(* IEC 61131-3 sources: volt/packages/volt-lsp-iec/test-corpus/awa-palletizer/Device/Plc Logic/Application/Library Manager/L_TB2P_TechModulesBasic, 108 files *)

(* ---- L_TB2P_ALLOWEDDIRECTION.dut ---- *)
TYPE L_TB2P_ALLOWEDDIRECTION :
(
	BOTH := 0,
	POSITIVE := 1,
	NEGATIVE := 2
);
END_TYPE

(* ---- L_TB2P_BASEIN.dut ---- *)
TYPE L_TB2P_BASEIN :
STRUCT
	XENABLE : BOOL;
	XRESETERROR : BOOL;
END_STRUCT
END_TYPE

(* ---- L_TB2P_BASEOUT.dut ---- *)
TYPE L_TB2P_BASEOUT :
STRUCT
	EERRORID : L_IE1P_Error;
	XWARNING : BOOL;
	XERROR : BOOL;
	ETMSTATE : L_TB2P_States := L_TB2P_States.DISABLED;
END_STRUCT
END_TYPE

(* ---- L_TB2P_BASICMOTIONBASEIN.dut ---- *)
TYPE L_TB2P_BASICMOTIONBASEIN :
STRUCT
	XUSEORIGINAL : BOOL;
	XENABLEOPERATION : BOOL;
	XQSPAPPLICATION : BOOL;
	XABORT : BOOL;
	XJOGPOS : BOOL;
	XJOGNEG : BOOL;
	XHOMEEXECUTE : BOOL;
	LROVERRIDE : LREAL := 1;
	SCCTRLBASICMOTION : L_TB2P_scCtrlBasicMotion;
END_STRUCT
END_TYPE

(* ---- L_TB2P_BASICMOTIONBASEOUT.dut ---- *)
TYPE L_TB2P_BASICMOTIONBASEOUT :
STRUCT
	XREADYFOROPERATION : BOOL;
	XOPERATIONENABLED : BOOL;
	XREADYFORMOTION : BOOL;
	XSTOACTIVE : BOOL;
	XQSPACTIVE : BOOL;
	XABORTBUSY : BOOL;
	XABORTDONE : BOOL;
	XJOGGINGBUSY : BOOL;
	XHOMINGBUSY : BOOL;
	XHOMINGDONE : BOOL;
	XISHOMED : BOOL;
	SCSTATUSBASICMOTION : L_TB2P_scStatusBasicMotion;
	LRSETACCOUT : LREAL;
	LRACTVEL : LREAL;
	LRSETVELOUT : LREAL;
	LRACTPOS : LREAL;
	LRSETPOSOUT : LREAL;
	LRACTFOLLOWINGERROR : LREAL;
END_STRUCT
END_TYPE

(* ---- L_TB2P_CATEGORY.dut ---- *)
TYPE L_TB2P_CATEGORY :
(
	DUMMY := 0
);
END_TYPE

(* ---- L_TB2P_CLASSID.dut ---- *)
TYPE L_TB2P_CLASSID :
(
	DUMMY := 0
);
END_TYPE

(* ---- L_TB2P_CLUTCHDIRECTION.dut ---- *)
TYPE L_TB2P_CLUTCHDIRECTION :
(
	MCNEGATIVEDIRECTION := -1,
	MCCURRENTDIRECTION := 0,
	MCPOSITIVEDIRECTION := 1
);
END_TYPE

(* ---- L_TB2P_CLUTCHMODE.dut ---- *)
TYPE L_TB2P_CLUTCHMODE :
(
	ABSOLUTE := 0,
	RELATIVE := 1,
	RAMP_POS := 2,
	RAMP_TIME := 3,
	DISTABSOLUTE := 4,
	ABSOLUTE_IN_TARGET := 5,
	DISTRELATIVE := 6,
	PROFGENABSOLUTE := 7,
	PROFGENRELATIVE := 8
);
END_TYPE

(* ---- L_TB2P_DIRECTION.dut ---- *)
TYPE L_TB2P_DIRECTION :
(
	BOTH := 0,
	DIRECTIONMASTER := 1
);
END_TYPE

(* ---- L_TB2P_ESELECTIONEXTTORQUELIMIT.dut ---- *)
TYPE L_TB2P_ESELECTIONEXTTORQUELIMIT :
(
	BOTHDIRECTIONS := 0,
	POSITIVEONLY := 1,
	NEGATIVEONLY := 2
);
END_TYPE

(* ---- L_TB2P_ESELECTIONMONITORINGSIGNALS.dut ---- *)
TYPE L_TB2P_ESELECTIONMONITORINGSIGNALS :
(
	NONE := 0,
	ACTUALMOTORTEMPERATURE := 1,
	ACTUALMOTORCURRENT := 2,
	DC_BUSVOLTAGE := 3,
	THERMALLOADDEVICE := 4,
	THERMALLOADMOTOR := 5,
	ANALOGSIGNAL := 6
);
END_TYPE

(* ---- L_TB2P_FBSTATES.dut ---- *)
TYPE L_TB2P_FBSTATES :
(
	INIT := 1,
	READY := 2,
	HOMING := 3,
	JOGGING := 10,
	JOGPOS := 11,
	JOGNEG := 12,
	POSITION_TRIMMING := 20,
	TRIM_POS_PLUS := 21,
	TRIM_POS_MINUS := 22,
	SYNCPOS := 30,
	POS_IS_SYNCHRONISED := 31,
	POSITIONING_TO_START_POS := 32,
	SYNCSPEED := 40,
	SPEED_IS_SYNCHRONISED := 41,
	DECOUPLED_LOCAL_DRIVING := 50,
	BASEVELOCITY := 51,
	CONTMOTION := 60,
	PREPARING_PATH := 61,
	CHECK_LIMITS := 62,
	SYNCLINEVEL := 70,
	CAMMING := 80,
	CAMMING_DONE := 81,
	CLUTCH_OPEN_INSTANT := 82,
	CLUTCH_CLOSE := 83,
	CLUTCH_OPEN := 84,
	CYCLICMOTION := 130,
	SETPARAMETERS := 140,
	CAMSEQUENCER_LOADCAMTABLE := 150,
	CAMSEQUENCER_CYCLICCAM1 := 151,
	CAMSEQUENCER_CYCLICCAM3 := 152,
	CAMSEQUENCER_CAM1CYCLICCAM3CAM1 := 153,
	CAMSEQUENCER_CAM1CAM2CYCLICCAM3CAM4CAM1 := 154,
	CALCULATION := 798,
	BUSY := 799,
	DONE := 800,
	EMERGENCYSTOP := 991,
	SLOWSTOP := 992,
	ABC := 993,
	STANDBY := 994,
	HALT := 995,
	STOP := 996,
	QUICKSTOP := 997,
	SERVICE := 998,
	ERROR := 999,
	SYSTEMFAULT := 1000
);
END_TYPE

(* ---- L_TB2P_INTERFACEID.dut ---- *)
TYPE L_TB2P_INTERFACEID :
(
	L_TB2P_ITECHMODULEBASE := (L_TB2P_Internal.cdiEnumStartValue + 1),
	L_TB2P_ITECHMODULEINTERNAL := (L_TB2P_Internal.cdiEnumStartValue + 2),
	L_TB2M_IERRORMANAGER := (L_TB2P_Internal.cdiEnumStartValue + 22),
	L_TB2P_ISTRUCTPROVIDER := (L_TB2P_Internal.cdiEnumStartValue + 23)
);
END_TYPE

(* ---- L_TB2P_SCAP_BASICMOTIONBASE.dut ---- *)
TYPE L_TB2P_SCAP_BASICMOTIONBASE :
STRUCT
END_STRUCT
END_TYPE

(* ---- L_TB2P_SCAP_TM_MOTIONCONTROL.dut ---- *)
TYPE L_TB2P_SCAP_TM_MOTIONCONTROL :
STRUCT
	AP_XDISABLEINTERNALCONTROL : BOOL;
END_STRUCT
END_TYPE

(* ---- L_TB2P_SCCTRLBASICMOTION.dut ---- *)
TYPE L_TB2P_SCCTRLBASICMOTION :
STRUCT
	XENABLEPOSITIVE : BOOL := TRUE;
	XENABLENEGATIVE : BOOL := TRUE;
	LROVERRIDEACC : LREAL := 1;
	LROVERRIDEJERK : LREAL := 1;
	XDISABLESWLIMIT : BOOL;
	XCONTINUOUSUPDATE : BOOL := TRUE;
	XHALT : BOOL;
	XFINISHPOSITIONING : BOOL;
	XMOVEVELEXECUTE : BOOL;
	XMOVEABSEXECUTE : BOOL;
	XMOVERELEXECUTE : BOOL;
	LRPOS_DIST : LREAL := 0;
	XHOMEABSSWITCH : BOOL;
	XRESETHOMEPOSITION : BOOL;
	XHWLIMITPOS : BOOL;
	XHWLIMITNEG : BOOL;
END_STRUCT
END_TYPE

(* ---- L_TB2P_SCCTRLBASICMOTIONEXTENDED.dut ---- *)
TYPE L_TB2P_SCCTRLBASICMOTIONEXTENDED :
STRUCT
	XENABLEOPERATION : BOOL;
	XRESETERROR : BOOL;
	XQSPAPPLICATION : BOOL;
	XABORT : BOOL;
	XJOGPOS : BOOL;
	XJOGNEG : BOOL;
	XHOMEEXECUTE : BOOL;
	LROVERRIDE : LREAL := 1;
	LRVEL : LREAL := 3600;
	LRACC : LREAL := 36000;
	LRDEC : LREAL := 36000;
	LRJERK : LREAL := 0;
	EDIRECTION : MC_DIRECTION := MC_DIRECTION.mcPositiveDirection;
	SCHOMEEXTTP : MC_TRIGGER_REF;
END_STRUCT
END_TYPE

(* ---- L_TB2P_SCDATABASICMOTIONBASE.dut ---- *)
TYPE L_TB2P_SCDATABASICMOTIONBASE :
STRUCT
	XHWLIMITSWITCH : BOOL;
	XENABLEOPERATION : BOOL;
	XHALT : BOOL;
	XABORT : BOOL;
	XHOMEEXECUTE : BOOL;
	XJOGPOS : BOOL;
	XJOGNEG : BOOL;
	XFINISHPOSITIONING : BOOL;
	XFINISHAVAILABLEMOVEABS : BOOL;
	XFINISHAVAILABLEMOVEREL : BOOL;
	XFINISHAVAILABLEMOVEVEL : BOOL;
	XMOVEVELEXECUTE : BOOL;
	XMOVEABSEXECUTE : BOOL;
	XMOVERELEXECUTE : BOOL;
	XRESETERROR : BOOL;
	XSPECIALABORTBEHAVIOR : BOOL;
	XSPECIALABORTBEHAVIORABC : BOOL;
	LRABORTDEC : LREAL;
	LRABORTJERK : LREAL;
	EFUNSTATEACT : L_MC1P_ABC_State;
	ECONTROLMODE : L_MC1P_ControlMode;
	XSTOACTIVE : BOOL;
	EAXISERRORID : L_IE1P_Error;
END_STRUCT
END_TYPE

(* ---- L_TB2P_SCPAR_BASICMOTIONBASE.dut ---- *)
TYPE L_TB2P_SCPAR_BASICMOTIONBASE :
STRUCT
END_STRUCT
END_TYPE

(* ---- L_TB2P_SCPAR_TM_MOTIONCONTROL.dut ---- *)
TYPE L_TB2P_SCPAR_TM_MOTIONCONTROL :
STRUCT
	LRVEL : LREAL := 3600;
	LRACC : LREAL := 36000;
	LRDEC : LREAL := 36000;
	LRJERK : LREAL := 0;
	EDIRECTION : MC_DIRECTION := MC_DIRECTION.mcPositiveDirection;
	SCHOMEEXTTP : MC_TRIGGER_REF;
END_STRUCT
END_TYPE

(* ---- L_TB2P_SCSF_BASICMOTIONBASE.dut ---- *)
TYPE L_TB2P_SCSF_BASICMOTIONBASE :
STRUCT
END_STRUCT
END_TYPE

(* ---- L_TB2P_SCSF_TM_MOTIONCONTROL.dut ---- *)
TYPE L_TB2P_SCSF_TM_MOTIONCONTROL :
STRUCT
	MP_XMULTICOREACTIVE : BOOL;
	MP_XINTERNALCONTROLACTIVE : BOOL;
	MP_IAXISTASKINDEX : INT;
	MP_ICALLTASKINDEX : INT;
END_STRUCT
END_TYPE

(* ---- L_TB2P_SCSTATUSBASICMOTION.dut ---- *)
TYPE L_TB2P_SCSTATUSBASICMOTION :
STRUCT
	XFUNBUSY : BOOL;
	XFUNDONE : BOOL;
	XFUNCOMMANDABORTED : BOOL;
	XHALTBUSY : BOOL;
	XHALTDONE : BOOL;
	ECONTROLMODE : L_MC1P_ControlMode;
	XHWLIMITSWITCHNEG : BOOL;
	XHWLIMITSWITCHPOS : BOOL;
	XSWLIMITENABLED : BOOL;
	XSWLIMITSWITCHNEG : BOOL;
	XSWLIMITSWITCHPOS : BOOL;
	EAXISTYPE : L_MC1P_DriveType;
	EAXISSTATE : L_MC1P_AXIS_STATE;
	XAXISWARNING : BOOL;
	XAXISERROR : BOOL;
	XDRIVEWARNING : BOOL;
	XDRIVEERROR : BOOL;
	DWDRIVEERRORID : DWORD;
	XCONSTANTVELOCITY : BOOL;
	XACCELERATING : BOOL;
	XDECELERATING : BOOL;
	XDIRECTIONPOSITIVE : BOOL;
	XDIRECTIONNEGATIVE : BOOL;
	XINPOSITION : BOOL;
	XAXISAVAILABLE : BOOL;
	XSTANDSTILLSETVELOCITY : BOOL;
	XSTANDSTILLACTVELOCITY : BOOL;
END_STRUCT
END_TYPE

(* ---- L_TB2P_SCSTATUSBASICMOTIONEXTENDED.dut ---- *)
TYPE L_TB2P_SCSTATUSBASICMOTIONEXTENDED :
STRUCT
	XREADYFOROPERATION : BOOL;
	XOPERATIONENABLED : BOOL;
	XREADYFORMOTION : BOOL;
	EAXISERRORID : L_IE1P_Error;
	XSTOACTIVE : BOOL;
	XQSPACTIVE : BOOL;
	XABORTBUSY : BOOL;
	XABORTDONE : BOOL;
	XJOGGINGBUSY : BOOL;
	XHOMINGBUSY : BOOL;
	XHOMINGDONE : BOOL;
	XISHOMED : BOOL;
	LRACTVEL : LREAL;
	LRSETVELOUT : LREAL;
	LRACTPOS : LREAL;
	LRSETPOSOUT : LREAL;
	LRACTFOLLOWINGERROR : LREAL;
END_STRUCT
END_TYPE

(* ---- L_TB2P_STATES.dut ---- *)
TYPE L_TB2P_STATES :
(
	DISABLED := -1,
	STANDBY := 0,
	STOP := 1,
	HOMING := 2,
	JOGGING := 3,
	MOVEVEL := 4,
	MOVEABS := 5,
	MOVEREL := 6,
	EXTERNAL := 7,
	ERROR := 8,
	FINISHPOSITIONING := 9,
	VELOCITYMODE := 15,
	ACC_DEC_SYNC := 30,
	SYNCHRONISED := 31,
	POSITIONING_TO_START_POS := 32,
	CAMMING := 33,
	POSITIONING_TO_TARGET_POS := 34,
	POSITIONING_TO_PARK_POS := 35,
	MOVE_TO_TARGET_POS := 36,
	POSITIONING := 38,
	POSITIONFOLLOWER := 41,
	VELOCITYFOLLOWER := 42,
	TORQUEFOLLOWER := 43,
	BASEVELOCITY := 51,
	ACC_DEC := 52,
	CONTMOTION := 60,
	LINEJOGGING := 65,
	SYNCLINEVEL := 70,
	VELOCITYMASTER := 71,
	IDENTMINERTIA := 80,
	IDENTDIAMETER := 81,
	IDENTFRICTION := 90,
	DANCERCTRL := 100,
	TENSIONCTRL := 110,
	PREPARING_PATH := 112,
	MOVE_PP := 114,
	CHECK_LIMITS := 115,
	TRANSFORMATION := 116,
	PATH_INTERRUPT := 117,
	MOVEELLIPTICAL := 118,
	WAITTIME := 119,
	PATH_HOLD := 120,
	SELECTMODECSV := 121,
	SELECTMODECST := 122,
	SELECTMODECSP := 123,
	CYCLICMOTION := 130,
	CUTTING := 170,
	IN_PARK_POS := 171,
	ASYNC_PHASE := 172,
	ENTRY_IN_SYNC_PAHSE := 173,
	EXIT_SYNC_PHASE := 175,
	HOLD_IN_PARK_POS := 176,
	START_CAM := 177,
	STOP_CAM := 178,
	WAIT_OF_NEXT_CUT := 179,
	STOP_IN_PARK_POS := 180,
	MOVE_XY := 186,
	MAINTENANCE := 187,
	BRAKE_TEST := 188,
	BRAKE_GRINDIN := 189,
	TRAVERSING := 190,
	SAW_IN_PROCESS := 200,
	MOVE_TO_PARK_POS := 210,
	REGULATION := 211,
	IDENTIFICATION := 212,
	CONTROL := 213,
	GROUPPAUSE := 300,
	MOVELINABS := 301,
	MOVELINREL := 302,
	MOVEDIRABS := 303,
	MOVEDIRREL := 304,
	CUTTING_DONE := 800,
	INIT := 900,
	SYSTEMFAULT := 1000,
	QUICKSTOP := 2018,
	HALT := 2019,
	ABORT := 2020,
	MANUALMODEJOG := 2001,
	SERVICE := 2003,
	GROUPSETPOS := 2010,
	GROUPABORT := 2015,
	GROUPHALT := 2016,
	JOBMODE := 2021,
	STOP_SAW := 20000,
	START_SAW := 20001,
	SAW_SYNCHRONIZED := 20003,
	SAW_SYNCHRONIZING := 20002,
	MOVE_TO_LOWER_LIMIT := 20006,
	WAITING_FOR_NEXT_CUT := 20007,
	MOVE_GAP := 20004,
	SYNC_OUT := 20005,
	X_MOVEABS := 3004,
	Y_MOVEABS := 3104,
	XY_MOVEREL := 3005,
	MAINTENANCE_JOGGING := 3003,
	STOP_VELOCITYMASTER := 4071,
	ABORT_VELOCITYFOLLOWER := 4042,
	HALT_FOLLOWER := 4043,
	ABORT_POSITIONFOLLOWER := 4044
);
END_TYPE

(* ---- L_TB2P_SYNCMODE.dut ---- *)
TYPE L_TB2P_SYNCMODE :
(
	PROFGENABSOLUTE := 0,
	PROFGENRELATIVE := 1,
	DISTABSOLUTE := 2,
	DISTRELATIVE := 3,
	CAMABSOLUTE := 4,
	INSTANTABSOLUTE := 10,
	INSTANTRELATIVE := 11
);
END_TYPE

(* ---- L_TB2P_CONSTANTS.gvl ---- *)
VAR_GLOBAL
	GC_DWCHECKIDTAPPETREF : DWORD := 16#DC34;
	GC_LREPSILON : LREAL := 1E-06;
	GC_POSITIVE_LIMIT_32BIT : LREAL := 2147483647;
	GC_NEGATIVE_LIMIT_32BIT : LREAL := -2147483647;
	GC_PI : LREAL := 3.1415926535897931;
END_VAR

(* ---- L_TB2P_INTERNAL.gvl ---- *)
VAR_GLOBAL
	CDIENUMSTARTVALUE : DINT := 20000;
END_VAR

(* ---- L_TB2M_IERRORMANAGER.itf ---- *)
INTERFACE L_TB2M_IERRORMANAGER
END_INTERFACE

METHOD GETERROR : BOOL
VAR_OUTPUT
	EERRORID : L_IE1P_Error;
END_VAR
END_METHOD

METHOD GETWARNING : BOOL
VAR_OUTPUT
	EERRORID : L_IE1P_Error;
END_VAR
END_METHOD

METHOD RESETREQUESTWARNING
END_METHOD

METHOD SETERROR
VAR_INPUT
	EERRORID : L_IE1P_Error;
	ESEVERITY : L_IE1P_SeverityLevel;
END_VAR
END_METHOD

METHOD SETERROREXTERNAL
VAR_INPUT
	XERROR : BOOL;
	EERRORID : L_IE1P_Error;
END_VAR
END_METHOD

METHOD SETREQUESTCONDITIONWARNING
VAR_IN_OUT
	ITFREQUEST : L_UBUP_IRequest;
END_VAR
END_METHOD

METHOD SETWARNING
VAR_INPUT
	EWARNINGID : L_IE1P_Error;
END_VAR
END_METHOD

METHOD SETWARNINGEXTERNAL
VAR_INPUT
	XWARNING : BOOL;
	EWARNINGID : L_IE1P_Error;
END_VAR
END_METHOD

(* ---- L_TB2M_IERRORMANAGERCALLBACK.itf ---- *)
INTERFACE L_TB2M_IERRORMANAGERCALLBACK
END_INTERFACE

METHOD ERRORSTATUSINFO
VAR_INPUT
	XERROR : BOOL;
	XWARNING : BOOL;
	EERRORID : L_IE1P_Error;
END_VAR
END_METHOD

(* ---- L_TB2M_IEXTENDEDTECHNOLOGIE.itf ---- *)
INTERFACE L_TB2M_IEXTENDEDTECHNOLOGIE
END_INTERFACE

METHOD EXTENDEDCALLFBS
VAR_INPUT
	ECASE : L_UBUP_StateHandleCase;
END_VAR
END_METHOD

METHOD EXTENDEDFINALIZECYCLE : BOOL
END_METHOD

METHOD EXTENDEDHANDLESTATE
VAR_INPUT
	ITFPARENT : L_UBUP_IStateClient;
	ITFSTATESERVER : L_UBUP_IStateServer;
	ISTATE : INT;
	ECASE : L_UBUP_StateHandleCase;
END_VAR
END_METHOD

METHOD EXTENDEDHANDLETRANSITION
VAR_INPUT
	ITFSTATESERVER : L_UBUP_IStateServer;
END_VAR
END_METHOD

METHOD EXTENDEDPREPARECYCLE
END_METHOD

METHOD EXTENDEDSTIMULATEREQUESTS
VAR_INPUT
	ECASE : L_UBUP_StateHandleCase;
END_VAR
END_METHOD

METHOD PREPARESTATECHANGE
END_METHOD

(* ---- L_TB2P_IBASICMOTIONBASE.itf ---- *)
INTERFACE L_TB2P_IBASICMOTIONBASE
END_INTERFACE

METHOD CALL_ABC
VAR_INPUT
	ITFTECHMODULE : L_TB2P_IBasicMotionBase;
	XQSPAPPLICATION : BOOL;
	XHALT : BOOL;
	XABORT : BOOL;
	XHOMEEXECUTE : BOOL;
	XJOGPOS : BOOL;
	XJOGNEG : BOOL;
	XFINISHPOSITIONING : BOOL;
	XMOVEVELEXECUTE : BOOL;
	XMOVEABSEXECUTE : BOOL;
	XMOVERELEXECUTE : BOOL;
	XENABLEOPERATION : BOOL;
	XRESETERROR : BOOL;
	XENABLEPOSITIVE : BOOL;
	XENABLENEGATIVE : BOOL;
	XDISABLESWLIMIT : BOOL;
	LROVERRIDE : LREAL;
	LROVERRIDEACC : LREAL;
	LROVERRIDEJERK : LREAL;
	XRESETHOMEPOSITION : BOOL;
	XCONTINUOUSUPDATE : BOOL;
	LRPOS_DIST : LREAL;
	LRVEL : LREAL;
	LRACC : LREAL;
	LRDEC : LREAL;
	LRJERK : LREAL;
	EDIRECTION : MC_DIRECTION;
	SCHOMEEXTTP : MC_TRIGGER_REF;
	XHOMEABSSWITCH : BOOL;
	XSPECIALABORTBEHAVIOR : BOOL;
	LRABORTDEC : LREAL;
	LRABORTJERK : LREAL;
END_VAR
VAR_OUTPUT
	XERROR : BOOL;
	EERRORID : L_IE1P_Error;
	XFUNBUSY : BOOL;
	XFUNDONE : BOOL;
	XFUNCOMMANDABORTED : BOOL;
	EFUNSTATEACT : L_MC1P_ABC_State;
	ECONTROLMODE : L_MC1P_ControlMode;
	XISHOMED : BOOL;
	XHWLIMITSWITCHNEG : BOOL;
	XHWLIMITSWITCHPOS : BOOL;
	XSWLIMITENABLED : BOOL;
	XSWLIMITSWITCHNEG : BOOL;
	XSWLIMITSWITCHPOS : BOOL;
	EAXISTYPE : L_MC1P_DriveType;
	EAXISSTATE : L_MC1P_AXIS_STATE;
	XSTOACTIVE : BOOL;
	XREADYFOROPERATION : BOOL;
	XOPERATIONENABLED : BOOL;
	XREADYFORMOTION : BOOL;
	XAXISWARNING : BOOL;
	XAXISERROR : BOOL;
	EAXISERRORID : L_IE1P_Error;
	XDRIVEWARNING : BOOL;
	XDRIVEERROR : BOOL;
	DWDRIVEERRORID : DWORD;
	LRACTPOS : LREAL;
	LRACTVEL : LREAL;
	LRSETPOSOUT : LREAL;
	LRSETVELOUT : LREAL;
	LRACTFOLLOWINGERROR : LREAL;
	XINPOSITION : BOOL;
	XSTANDSTILLSETVELOCITY : BOOL;
	XSTANDSTILLACTVELOCITY : BOOL;
	XCONSTANTVELOCITY : BOOL;
	XACCELERATING : BOOL;
	XDECELERATING : BOOL;
	XDIRECTIONPOSITIVE : BOOL;
	XDIRECTIONNEGATIVE : BOOL;
	XAXISAVAILABLE : BOOL;
END_VAR
VAR_IN_OUT
	AXIS : AXIS_REF;
END_VAR
END_METHOD

(* ---- L_TB2P_ICONNECTORBASICMOTIONBASE.itf ---- *)
INTERFACE L_TB2P_ICONNECTORBASICMOTIONBASE
END_INTERFACE

(* ---- L_TB2P_ISTRUCTPROVIDER.itf ---- *)
INTERFACE L_TB2P_ISTRUCTPROVIDER
END_INTERFACE

METHOD GET_PAP : POINTER TO L_TB2P_scAP_TM_MotionControl
END_METHOD

METHOD GET_PPAR : POINTER TO L_TB2P_scPar_TM_MotionControl
END_METHOD

METHOD GET_PSF : POINTER TO L_TB2P_scSF_TM_MotionControl
END_METHOD

(* ---- L_TB2P_ITECHMODULEBASE.itf ---- *)
INTERFACE L_TB2P_ITECHMODULEBASE
END_INTERFACE

(* ---- L_TB2P_ITECHMODULEINTERNAL.itf ---- *)
INTERFACE L_TB2P_ITECHMODULEINTERNAL
END_INTERFACE

METHOD HANDOVERRESOURCE : BOOL
VAR_INPUT
	ITFRESOURCE : L_UBUP_IUnknown;
END_VAR
END_METHOD

(* ---- L_TB2P_ITM_BASE.itf ---- *)
INTERFACE L_TB2P_ITM_BASE
END_INTERFACE

METHOD SETADDMODULEINFO
VAR_INPUT
	ESUBCOMPTYPE : UDINT;
	SLICINFO : STRING(10);
END_VAR
END_METHOD

(* ---- GETBOOLEANPROPERTY.pou ---- *)
FUNCTION GETBOOLEANPROPERTY : BOOL
VAR_INPUT
	STKEY : WSTRING;
END_VAR
END_FUNCTION

(* ---- GETCOMPANY.pou ---- *)
FUNCTION GETCOMPANY : WSTRING
END_FUNCTION

(* ---- GETNUMBERPROPERTY.pou ---- *)
FUNCTION GETNUMBERPROPERTY : DINT
VAR_INPUT
	STKEY : WSTRING;
END_VAR
END_FUNCTION

(* ---- GETTEXTPROPERTY.pou ---- *)
FUNCTION GETTEXTPROPERTY : WSTRING
VAR_INPUT
	STKEY : WSTRING;
END_VAR
END_FUNCTION

(* ---- GETTEXTPROPERTY2.pou ---- *)
FUNCTION GETTEXTPROPERTY2 : POINTER TO WSTRING
VAR_INPUT
	STKEY : WSTRING;
END_VAR
END_FUNCTION

(* ---- GETTITLE.pou ---- *)
FUNCTION GETTITLE : WSTRING
END_FUNCTION

(* ---- GETVERSION.pou ---- *)
FUNCTION GETVERSION : VERSION
END_FUNCTION

(* ---- GETVERSIONPROPERTY.pou ---- *)
FUNCTION GETVERSIONPROPERTY : VERSION
VAR_INPUT
	STKEY : WSTRING;
END_VAR
END_FUNCTION

(* ---- L_TB2P_CONVERTPOSTOMODULOPOS.pou ---- *)
FUNCTION L_TB2P_CONVERTPOSTOMODULOPOS : LREAL
VAR_INPUT
	LRPOS : LREAL;
	LRPERIOD : LREAL;
END_VAR
VAR_OUTPUT
	DIREVCOUNTER : DINT;
END_VAR
END_FUNCTION

(* ---- L_TB2P_CONVERTPOSTOMODULOPOSEXTENDED.pou ---- *)
FUNCTION L_TB2P_CONVERTPOSTOMODULOPOSEXTENDED : LREAL
VAR_INPUT
	LRPOS : LREAL;
	LRPERIOD : LREAL;
END_VAR
VAR_OUTPUT
	DIREVCOUNTER : DINT;
END_VAR
END_FUNCTION

(* ---- L_TB2P_HLPCALCTARGETANDKOEFPOLY5THORD.pou ---- *)
FUNCTION L_TB2P_HLPCALCTARGETANDKOEFPOLY5THORD : ARRAY [0..5] OF LREAL
VAR_INPUT
	LRYVELSTART : LREAL;
	LRYVELEND : LREAL;
END_VAR
VAR_OUTPUT
	ALRKOEF : ARRAY [0..5] OF LREAL;
	LRYPOSEND : LREAL;
END_VAR
END_FUNCTION

(* ---- L_TB2P_HLPCALCYOFPOLY5THORDBASE.pou ---- *)
FUNCTION L_TB2P_HLPCALCYOFPOLY5THORDBASE : LREAL
VAR_OUTPUT
	LRYPOSSCALED : LREAL;
END_VAR
VAR_IN_OUT
	LRXPOSSCALED : LREAL;
	ALRKOEF : ARRAY [0..5] OF LREAL;
END_VAR
END_FUNCTION

(* ---- L_TB2P_HLPDELTAVELTIMEEXTENDED.pou ---- *)
FUNCTION L_TB2P_HLPDELTAVELTIMEEXTENDED : BOOL
VAR_INPUT
	LRVELSTART : LREAL;
	LRACCSTART : LREAL;
	LRMAXACC : LREAL;
	LRMAXJERK : LREAL;
END_VAR
VAR_OUTPUT
	LRTIME : LREAL;
	LRDIST : LREAL;
END_VAR
END_FUNCTION

(* ---- L_TB2P_HLPDELTAVELTIMETOCONTANTVEL.pou ---- *)
FUNCTION L_TB2P_HLPDELTAVELTIMETOCONTANTVEL : BOOL
VAR_INPUT
	LRACCSTART : LREAL;
	LRMAXJERK : LREAL;
	WMODE : WORD;
END_VAR
VAR_OUTPUT
	LRVEL : LREAL;
	LRTIME : LREAL;
	LRDIST : LREAL;
END_VAR
END_FUNCTION

(* ---- L_TB2P_HLPMODULODIFF.pou ---- *)
FUNCTION L_TB2P_HLPMODULODIFF : LREAL
VAR_INPUT
	LRDIFF : LREAL;
	LRLEN : LREAL;
END_VAR
END_FUNCTION

(* ---- L_TB2P_HLPTIMEMOVEDIST.pou ---- *)
FUNCTION L_TB2P_HLPTIMEMOVEDIST : BOOL
VAR_INPUT
	LRDIST : LREAL;
	LRVEL : LREAL;
	LRACC : LREAL;
END_VAR
VAR_OUTPUT
	LRTIME : LREAL;
END_VAR
END_FUNCTION

(* ---- L_TB2P_LREQ.pou ---- *)
FUNCTION L_TB2P_LREQ : BOOL
VAR_INPUT
	LRVALUE : LREAL;
	LRTARGET : LREAL;
END_VAR
END_FUNCTION

(* ---- L_TB2P_LRGE.pou ---- *)
FUNCTION L_TB2P_LRGE : BOOL
VAR_INPUT
	LRVALUE : LREAL;
	LRTARGET : LREAL;
END_VAR
END_FUNCTION

(* ---- L_TB2P_LRGT.pou ---- *)
FUNCTION L_TB2P_LRGT : BOOL
VAR_INPUT
	LRVALUE : LREAL;
	LRTARGET : LREAL;
END_VAR
END_FUNCTION

(* ---- L_TB2P_LRLE.pou ---- *)
FUNCTION L_TB2P_LRLE : BOOL
VAR_INPUT
	LRVALUE : LREAL;
	LRTARGET : LREAL;
END_VAR
END_FUNCTION

(* ---- L_TB2P_LRLT.pou ---- *)
FUNCTION L_TB2P_LRLT : BOOL
VAR_INPUT
	LRVALUE : LREAL;
	LRTARGET : LREAL;
END_VAR
END_FUNCTION

(* ---- L_TB2P_LRNE.pou ---- *)
FUNCTION L_TB2P_LRNE : BOOL
VAR_INPUT
	LRVALUE : LREAL;
	LRTARGET : LREAL;
END_VAR
END_FUNCTION

(* ---- L_TB2P_TRANSITIONBASEVEL.pou ---- *)
FUNCTION L_TB2P_TRANSITIONBASEVEL : BOOL
VAR_INPUT
	LRSETBASEVEL : LREAL;
	XRTRIGSETBASEVEL : BOOL;
	XSYNCIN : BOOL;
	XJOGPOS : BOOL;
	XJOGNEG : BOOL;
	XQSPAPPLICATION : BOOL;
	XHALT : BOOL;
	XABORT : BOOL;
	EACTTMSTATE : L_TB2P_States;
	DWLIMITERCONTROL : DWORD;
	EALLOWEDDIRECTION : L_TB2P_AllowedDirection;
END_VAR
VAR_OUTPUT
	XDIRECTIONDISABLED : BOOL;
END_VAR
VAR_IN_OUT
	AXIS : AXIS_REF;
END_VAR
END_FUNCTION

(* ---- L_TB2P_TRANSITIONJOGGING.pou ---- *)
FUNCTION L_TB2P_TRANSITIONJOGGING : BOOL
VAR_INPUT
	XRTRIGJOGPOS : BOOL;
	XRTRIGJOGNEG : BOOL;
	XJOGPOS : BOOL;
	XJOGNEG : BOOL;
	XQSPAPPLICATION : BOOL;
	XHALT : BOOL;
	XABORT : BOOL;
	EACTTMSTATE : L_TB2P_States;
	DWLIMITERCONTROL : DWORD;
	EALLOWEDDIRECTION : L_TB2P_AllowedDirection;
END_VAR
VAR_OUTPUT
	XDIRECTIONDISABLED : BOOL;
END_VAR
VAR_IN_OUT
	AXIS : AXIS_REF;
END_VAR
END_FUNCTION

(* ---- L_TB2P_TRANSITIONLEVELFUN.pou ---- *)
FUNCTION L_TB2P_TRANSITIONLEVELFUN : BOOL
VAR_INPUT
	XRTRIGFUN : BOOL;
	XFUNCTION : BOOL;
	XJOGPOS : BOOL;
	XJOGNEG : BOOL;
	XQSPAPPLICATION : BOOL;
	XBLOCKFUN1 : BOOL;
	XBLOCKFUN2 : BOOL;
	XBLOCKFUN3 : BOOL;
	XBLOCKFUN4 : BOOL;
	EACTTMSTATE : L_TB2P_States;
	EALLOWEDTMSTATE1 : L_TB2P_States := L_TB2P_States.STANDBY;
	EALLOWEDTMSTATE2 : L_TB2P_States := L_TB2P_States.STANDBY;
	EALLOWEDTMSTATE3 : L_TB2P_States := L_TB2P_States.STANDBY;
	EALLOWEDTMSTATE4 : L_TB2P_States := L_TB2P_States.STANDBY;
	EBLOCKTMSTATE1 : L_TB2P_States := L_TB2P_States.DISABLED;
	EBLOCKTMSTATE2 : L_TB2P_States := L_TB2P_States.DISABLED;
	DWLIMITERCONTROL : DWORD;
END_VAR
VAR_IN_OUT
	AXIS : AXIS_REF;
END_VAR
END_FUNCTION

(* ---- L_TB2P_TRANSITIONMOVEPROFILE.pou ---- *)
FUNCTION L_TB2P_TRANSITIONMOVEPROFILE : BOOL
VAR_INPUT
	XRTRIGMOVEPROFILE : BOOL;
	XMOVEPROFILE : BOOL;
	IPROFILEDIRECTION : INT := 0;
	XJOGPOS : BOOL;
	XJOGNEG : BOOL;
	XQSPAPPLICATION : BOOL;
	EACTTMSTATE : L_TB2P_States;
	DWLIMITERCONTROL : DWORD;
	EALLOWEDDIRECTION : L_TB2P_AllowedDirection;
END_VAR
VAR_OUTPUT
	XDIRECTIONDISABLED : BOOL;
END_VAR
VAR_IN_OUT
	AXIS : AXIS_REF;
END_VAR
END_FUNCTION

(* ---- L_TB2P_TRANSITIONSYNCIN.pou ---- *)
FUNCTION L_TB2P_TRANSITIONSYNCIN : BOOL
VAR_INPUT
	XRTRIGSYNCIN : BOOL;
	XSYNCIN : BOOL;
	XJOGPOS : BOOL;
	XJOGNEG : BOOL;
	XQSPAPPLICATION : BOOL;
	EACTTMSTATE : L_TB2P_States;
	DWLIMITERCONTROL : DWORD;
END_VAR
VAR_IN_OUT
	AXIS : AXIS_REF;
END_VAR
END_FUNCTION

(* ---- L_TB2P_TRANSITIONSYNCINALLOWEDDIRECTION.pou ---- *)
FUNCTION L_TB2P_TRANSITIONSYNCINALLOWEDDIRECTION : BOOL
VAR_INPUT
	XACTMASTERDIRVALID : BOOL;
	IACTMASTERDIRECTION : INT := 0;
	LRCYCLELENGTH : LREAL;
	LRMASTERPOSFORSYNC : LREAL;
	LRSETSLAVEPOS : LREAL;
	LRMASTERVELFORSYNC : LREAL;
	LRSETSLAVEVELOCITY : LREAL;
	DWLIMITERCONTROL : DWORD;
	EALLOWEDDIRECTION : L_TB2P_AllowedDirection;
	ESYNCMODE : L_TB2P_SyncMode;
	LRSYNCVEL : LREAL;
	LRSLAVESYNCINDIST : LREAL;
END_VAR
VAR_OUTPUT
	XINVALIDMASTERDIRECTION : BOOL;
	XDIRECTIONDISABLED : BOOL;
END_VAR
VAR_IN_OUT
	AXIS : AXIS_REF;
END_VAR
END_FUNCTION

(* ---- GLOBALTEXTLIST.pou ---- *)
FUNCTION_BLOCK GLOBALTEXTLIST
VAR
	M_TEXTLISTFILE : STRING(255);
	_STNAMESPACE : STRING;
END_VAR
END_FUNCTION_BLOCK

(* ---- L_TB2M_BASICMOTIONBASE.pou ---- *)
FUNCTION_BLOCK L_TB2M_BASICMOTIONBASE EXTENDS L_TB2P_TechModuleBase
VAR_INPUT
	XUSEORIGINAL : BOOL;
	XENABLE : BOOL;
	XENABLEOPERATION : BOOL;
	XRESETERROR : BOOL;
	XQSPAPPLICATION : BOOL;
	XABORT : BOOL;
	XJOGPOS : BOOL;
	XJOGNEG : BOOL;
	XHOMEEXECUTE : BOOL;
	LROVERRIDE : LREAL := 1;
	SCCTRLBASICMOTION : L_TB2P_scCtrlBasicMotion;
	SCPAR : L_TB2P_scPar_BasicMotionBase;
	SCACCESSPOINTS : L_TB2P_scAP_BasicMotionBase;
END_VAR
VAR_OUTPUT
	XREADYFOROPERATION : BOOL;
	XOPERATIONENABLED : BOOL;
	XREADYFORMOTION : BOOL;
	XERROR : BOOL;
	XWARNING : BOOL;
	EERRORID : L_IE1P_Error;
	XSTOACTIVE : BOOL;
	XQSPACTIVE : BOOL;
	XABORTBUSY : BOOL;
	XABORTDONE : BOOL;
	XJOGGINGBUSY : BOOL;
	XHOMINGBUSY : BOOL;
	XHOMINGDONE : BOOL;
	XISHOMED : BOOL;
	ETMSTATE : L_TB2P_States := L_TB2P_States.DISABLED;
	SCSTATUSBASICMOTION : L_TB2P_scStatusBasicMotion;
	LRSETACCOUT : LREAL;
	LRACTVEL : LREAL;
	LRSETVELOUT : LREAL;
	LRACTPOS : LREAL;
	LRSETPOSOUT : LREAL;
	LRACTFOLLOWINGERROR : LREAL;
	SCSIGNALFLOW : L_TB2P_scSF_BasicMotionBase;
END_VAR
VAR_IN_OUT
	AXIS : AXIS_REF;
END_VAR
VAR
	XUSEORIGINAL_OLD : BOOL;
	TM_INT : L_TB2M_TM_MotionControl;
	SCPAR_INT : L_TB2P_scPar_BasicMotionBase;
	_UICALLMFUNIDXINPUT : UINT := 1;
	_UICALLMFUNIDXOUTPUT : UINT := 1;
	_ASCINPUT : ARRAY [1.._MCCall.c_BufferDepthInput] OF L_TB2P_BasicMotionBaseIn;
	_ASCOUTPUT : ARRAY [1.._MCCall.c_BufferDepthOutput] OF L_TB2P_BasicMotionBaseOut;
	_ASCPARCORE : ARRAY [1.._MCCall.c_BufferDepthInput] OF L_TB2P_scPar_BasicMotionBase;
	_ASCAP : ARRAY [1.._MCCall.c_BufferDepthInput] OF L_TB2P_scAP_BasicMotionBase;
	_ASCSF : ARRAY [1.._MCCall.c_BufferDepthOutput] OF L_TB2P_scSF_BasicMotionBase;
	_SCACCESSPOINTSCORE : L_TB2P_scAP_BasicMotionBase;
	_SCSIGNALFLOWCORE : L_TB2P_scSF_BasicMotionBase;
	_MCCALL : L_UM1P_MCCall;
	_SCINPUTVISU : L_TB2P_BasicMotionBaseIn;
	_PSCINPUTVISU : POINTER TO L_TB2P_BasicMotionBaseIn := ADR(_scInputVisu);
	_PSCOUTPUTVISU : POINTER TO L_TB2P_BasicMotionBaseOut := ADR(_ascOutput[1]);
	_PSCPARVISU : POINTER TO L_TB2P_scPar_BasicMotionBase := ADR(scPar_int);
	DECORATOR : L_UBUP_IStateClientDecorator;
	ITFBASICMOTION : L_TB2P_IBasicMotionBase;
	ITFITECHMODULEINTERNAL : L_TB2P_ITechModuleInternal;
	LRJERKDEC : LREAL;
	LRJOGGINGJERKDEC : LREAL;
	MONITORSTATESERVER : L_UBUP_IMonitorStateServer;
	REMAININGTIMEOFPROFILE : LREAL;
	REMAININGTIMEOFPROFILEAVAILABLE : BOOL;
	STATESERVER : L_UBUP_IStateServer;
END_VAR
END_FUNCTION_BLOCK

METHOD CALL_ABC
VAR_INPUT
	ITFTECHMODULE : L_TB2P_IBasicMotionBase;
	XQSPAPPLICATION : BOOL;
	XHALT : BOOL;
	XABORT : BOOL;
	XHOMEEXECUTE : BOOL;
	XJOGPOS : BOOL;
	XJOGNEG : BOOL;
	XFINISHPOSITIONING : BOOL;
	XMOVEVELEXECUTE : BOOL;
	XMOVEABSEXECUTE : BOOL;
	XMOVERELEXECUTE : BOOL;
	XENABLEOPERATION : BOOL;
	XRESETERROR : BOOL;
	XENABLEPOSITIVE : BOOL;
	XENABLENEGATIVE : BOOL;
	XDISABLESWLIMIT : BOOL;
	LROVERRIDE : LREAL;
	LROVERRIDEACC : LREAL;
	LROVERRIDEJERK : LREAL;
	XRESETHOMEPOSITION : BOOL;
	XCONTINUOUSUPDATE : BOOL;
	LRPOS_DIST : LREAL;
	LRVEL : LREAL;
	LRACC : LREAL;
	LRDEC : LREAL;
	LRJERK : LREAL;
	EDIRECTION : MC_DIRECTION;
	SCHOMEEXTTP : MC_TRIGGER_REF;
	XHOMEABSSWITCH : BOOL;
	XSPECIALABORTBEHAVIOR : BOOL;
	LRABORTDEC : LREAL;
	LRABORTJERK : LREAL;
END_VAR
VAR_OUTPUT
	XERROR : BOOL;
	EERRORID : L_IE1P_Error;
	XFUNBUSY : BOOL;
	XFUNDONE : BOOL;
	XFUNCOMMANDABORTED : BOOL;
	EFUNSTATEACT : L_MC1P_ABC_State;
	ECONTROLMODE : L_MC1P_ControlMode;
	XISHOMED : BOOL;
	XHWLIMITSWITCHNEG : BOOL;
	XHWLIMITSWITCHPOS : BOOL;
	XSWLIMITENABLED : BOOL;
	XSWLIMITSWITCHNEG : BOOL;
	XSWLIMITSWITCHPOS : BOOL;
	EAXISTYPE : L_MC1P_DriveType;
	EAXISSTATE : L_MC1P_AXIS_STATE;
	XSTOACTIVE : BOOL;
	XREADYFOROPERATION : BOOL;
	XOPERATIONENABLED : BOOL;
	XREADYFORMOTION : BOOL;
	XAXISWARNING : BOOL;
	XAXISERROR : BOOL;
	EAXISERRORID : L_IE1P_Error;
	XDRIVEWARNING : BOOL;
	XDRIVEERROR : BOOL;
	DWDRIVEERRORID : DWORD;
	LRACTPOS : LREAL;
	LRACTVEL : LREAL;
	LRSETPOSOUT : LREAL;
	LRSETVELOUT : LREAL;
	LRACTFOLLOWINGERROR : LREAL;
	XINPOSITION : BOOL;
	XSTANDSTILLSETVELOCITY : BOOL;
	XSTANDSTILLACTVELOCITY : BOOL;
	XCONSTANTVELOCITY : BOOL;
	XACCELERATING : BOOL;
	XDECELERATING : BOOL;
	XDIRECTIONPOSITIVE : BOOL;
	XDIRECTIONNEGATIVE : BOOL;
	XAXISAVAILABLE : BOOL;
END_VAR
VAR_IN_OUT
	AXIS : AXIS_REF;
END_VAR
END_METHOD

METHOD CALL_HWLIMITSWITCH
VAR_INPUT
	ITFTECHMODULE : L_TB2P_IBasicMotionBase;
	XENABLE : BOOL;
	XLIMITSWITCHPOS : BOOL;
	XLIMITSWITCHNEG : BOOL;
END_VAR
VAR_OUTPUT
	XBUSY : BOOL;
	XERROR : BOOL;
	EERRORID : L_IE1P_Error;
END_VAR
END_METHOD

METHOD GET_PAP : POINTER TO L_TB2P_scAP_TM_MotionControl
END_METHOD

METHOD GET_PPAR : POINTER TO L_TB2P_scPar_TM_MotionControl
END_METHOD

METHOD GET_PSF : POINTER TO L_TB2P_scSF_TM_MotionControl
END_METHOD

METHOD CALLFUNCTION
VAR_INPUT
	UIINPUTDATAIDX : UINT;
	UIOUTPUTDATAIDX : UINT;
END_VAR
END_METHOD

METHOD COPYINPUTS : BOOL
VAR_INPUT
	IDX : WORD;
END_VAR
END_METHOD

METHOD COPYOUTPUTS : BOOL
VAR_INPUT
	IDX : WORD;
END_VAR
END_METHOD

METHOD FUNCTIONWASCALLEDTWICE : BOOL
VAR_INPUT
	IDX : WORD;
END_VAR
END_METHOD

METHOD HANDLESTANDARDCALL : BOOL
END_METHOD

METHOD SYNCOUTPUTS
VAR_INPUT
	UICOPYOUTPUTFROMIDX : UINT;
	UICOPYOUTPUTTOIDX : UINT;
END_VAR
END_METHOD

METHOD FB_INIT : BOOL
VAR_INPUT
	BINITRETAINS : BOOL;
	BINCOPYCODE : BOOL;
END_VAR
END_METHOD

METHOD CALL_INTERNALCTRL
END_METHOD

METHOD SETERROR
VAR_INPUT
	XERROR : BOOL;
	EERRORID : L_IE1P_Error;
END_VAR
END_METHOD

(* ---- L_TB2M_ERRORMANAGER.pou ---- *)
FUNCTION_BLOCK L_TB2M_ERRORMANAGER EXTENDS L_TB2M_ErrorManagerBase
VAR_INPUT
	ERRORHANDLER : L_IE1P_IErrorHandler;
END_VAR
VAR
	_MODULEHANDLER : L_IMHP_IModuleHandler;
	FB_SETERROR : L_IE1P_SetError;
	FB_RESETERROR : L_IE1P_ResetError;
END_VAR
END_FUNCTION_BLOCK

METHOD INITIALIZE : BOOL
VAR_INPUT
	MODULEHANDLER : L_IMHP_IModuleHandler;
	ITFERRORMANAGERCALLBACK : L_TB2M_IErrorManagerCallback;
END_VAR
END_METHOD

METHOD DETECTERRORRESET : BOOL
VAR_INPUT
	XRESETERROR : BOOL;
END_VAR
END_METHOD

METHOD FORWARDERROR
VAR_INPUT
	XERROR : BOOL;
	EERRORID : L_IE1P_Error;
	ESEVERITY : L_IE1P_SeverityLevel;
END_VAR
END_METHOD

METHOD FORWARDWARNING
VAR_INPUT
	XWARNING : BOOL;
	EWARNINGID : L_IE1P_Error;
END_VAR
END_METHOD

(* ---- L_TB2M_ERRORMANAGERBASE.pou ---- *)
FUNCTION_BLOCK L_TB2M_ERRORMANAGERBASE
VAR_INPUT
	XENABLE : BOOL;
END_VAR
VAR_OUTPUT
	XTRIGGERRESETERRORACTIVE : BOOL;
END_VAR
VAR
	XERROR_INT : BOOL;
	XWARNING_INT : BOOL;
	EERRORID_INT : L_IE1P_Error;
	ACTWARNINGSTATUS : DWORD;
	ACTERRORSTATUS : DWORD;
	XRESETERROROLD : BOOL;
	_ITFREQUESTCONDITIONWARNING : L_UBUP_IRequest := 0;
	_ITFERRORMANAGERCALLBACK : L_TB2M_IErrorManagerCallback;
	C_MODWARNING : DWORD := 3;
	C_EXTWARNING : DWORD := 2;
	C_CONDWARNING : DWORD := 1;
	C_NOWARNING : DWORD := 0;
	C_MODERROR : DWORD := 3;
	C_EXTERROR : DWORD := 2;
	C_NOERROR : DWORD := 0;
END_VAR
END_FUNCTION_BLOCK

METHOD INITIALIZE : BOOL
VAR_INPUT
	MODULEHANDLER : L_IMHP_IModuleHandler;
	ITFERRORMANAGERCALLBACK : L_TB2M_IErrorManagerCallback;
END_VAR
END_METHOD

METHOD RESET : BOOL
VAR_INPUT
	XRESETERROR : BOOL;
END_VAR
END_METHOD

METHOD SETWARNINGSTATUS : BOOL
VAR_INPUT
	NEWWARNINGSTATUS : DWORD;
	EWARNINGID : L_IE1P_Error;
END_VAR
END_METHOD

METHOD UPDATECONDITIONWARNING
END_METHOD

METHOD UPDATESTATUSINFO
END_METHOD

METHOD DETECTERRORRESET : BOOL
VAR_INPUT
	XRESETERROR : BOOL;
END_VAR
END_METHOD

METHOD FORWARDERROR
VAR_INPUT
	XERROR : BOOL;
	EERRORID : L_IE1P_Error;
	ESEVERITY : L_IE1P_SeverityLevel;
END_VAR
END_METHOD

METHOD FORWARDWARNING
VAR_INPUT
	XWARNING : BOOL;
	EWARNINGID : L_IE1P_Error;
END_VAR
END_METHOD

METHOD GETERROR : BOOL
VAR_OUTPUT
	EERRORID : L_IE1P_Error;
END_VAR
END_METHOD

METHOD GETWARNING : BOOL
VAR_OUTPUT
	EERRORID : L_IE1P.L_IE1P_Error;
END_VAR
END_METHOD

METHOD RESETREQUESTWARNING
END_METHOD

METHOD SETERROR
VAR_INPUT
	EERRORID : L_IE1P_Error;
	ESEVERITY : L_IE1P_SeverityLevel;
END_VAR
END_METHOD

METHOD SETERROREXTERNAL
VAR_INPUT
	XERROR : BOOL;
	EERRORID : L_IE1P_Error;
END_VAR
END_METHOD

METHOD SETREQUESTCONDITIONWARNING
VAR_IN_OUT
	ITFREQUEST : L_UBUP_IRequest;
END_VAR
END_METHOD

METHOD SETWARNING
VAR_INPUT
	EWARNINGID : L_IE1P_Error;
END_VAR
END_METHOD

METHOD SETWARNINGEXTERNAL
VAR_INPUT
	XWARNING : BOOL;
	EWARNINGID : L_IE1P_Error;
END_VAR
END_METHOD

METHOD REQUESTINTERFACE : BOOL
VAR_INPUT
	ID : DINT;
	PITFUNKNOWN : POINTER TO L_UBUP_IUnknown;
END_VAR
END_METHOD

(* ---- L_TB2M_ERRORMANAGERFM.pou ---- *)
FUNCTION_BLOCK L_TB2M_ERRORMANAGERFM
VAR_INPUT
	XENABLE : BOOL;
END_VAR
VAR_OUTPUT
	XTRIGGERRESETERRORACTIVE : BOOL;
END_VAR
VAR
	XERROR : REFERENCE TO BOOL;
	XWARNING : REFERENCE TO BOOL;
	EERRORID : REFERENCE TO L_IE1P_Error;
	XERROR_INT : BOOL;
	XWARNING_INT : BOOL;
	EERRORID_INT : L_IE1P_Error;
	XEXTERNALWARNING : BOOL;
	XEXTERNALERROR : BOOL;
	XERROR_FIRST : BOOL;
	XRESETERROROLD : BOOL;
	_ITFREQUESTCONDITIONWARNING : L_UBUP_IRequest := 0;
	_XCONDITIONWARNING : BOOL;
	_ECONDITIONWARNINGID : L_IE1P_Error;
END_VAR
END_FUNCTION_BLOCK

METHOD INITIALIZE : BOOL
VAR_INPUT
	PXERROR : POINTER TO BOOL;
	PXWARNING : POINTER TO BOOL;
	PEERRORID : POINTER TO L_IE1P_Error;
END_VAR
END_METHOD

METHOD RESET : BOOL
VAR_INPUT
	XRESETERROR : BOOL;
END_VAR
END_METHOD

METHOD RESETWARNING : BOOL
VAR_INPUT
	EWARNINGID : L_IE1P_Error;
END_VAR
END_METHOD

METHOD UPDATESTATUSINFO
END_METHOD

METHOD GETERROR : BOOL
VAR_OUTPUT
	EERRORID : L_IE1P_Error;
END_VAR
END_METHOD

METHOD GETWARNING : BOOL
VAR_OUTPUT
	EERRORID : L_IE1P.L_IE1P_Error;
END_VAR
END_METHOD

METHOD RESETREQUESTWARNING
END_METHOD

METHOD SETERROR
VAR_INPUT
	EERRORID : L_IE1P_Error;
	ESEVERITY : L_IE1P_SeverityLevel;
END_VAR
END_METHOD

METHOD SETERROREXTERNAL
VAR_INPUT
	XERROR : BOOL;
	EERRORID : L_IE1P_Error;
END_VAR
END_METHOD

METHOD SETREQUESTCONDITIONWARNING
VAR_IN_OUT
	ITFREQUEST : L_UBUP_IRequest;
END_VAR
END_METHOD

METHOD SETWARNING
VAR_INPUT
	EWARNINGID : L_IE1P_Error;
END_VAR
END_METHOD

METHOD SETWARNINGEXTERNAL
VAR_INPUT
	XWARNING : BOOL;
	EWARNINGID : L_IE1P_Error;
END_VAR
END_METHOD

METHOD REQUESTINTERFACE : BOOL
VAR_INPUT
	ID : DINT;
	PITFUNKNOWN : POINTER TO L_UBUP_IUnknown;
END_VAR
END_METHOD

(* ---- L_TB2M_FM_BASE.pou ---- *)
FUNCTION_BLOCK L_TB2M_FM_BASE
VAR_INPUT
	XENABLE : BOOL;
END_VAR
VAR_OUTPUT
	EERRORID : L_IE1P_Error;
	XWARNING : BOOL;
	XERROR : BOOL;
END_VAR
VAR
	FB_STATESERVER : L_UBUP_StateServer := STRUCT(iFreezeRequestPrio := 10);
	FB_ERRORMANAGER_INT : L_TB2M_ErrorManagerFM;
	ITFERRORMANAGER : L_TB2M_IErrorManager := fB_ErrorManager_int;
	FB_TRANSITION2STANDBY : L_UBUP_RequestTransitionEdge;
	ERRORMANAGER : L_TB2M_IErrorManager;
END_VAR
END_FUNCTION_BLOCK

METHOD CALLFBS
VAR_INPUT
	ECASE : L_UBUP.L_UBUP_StateHandleCase;
END_VAR
END_METHOD

METHOD CALLSTATE
VAR_INPUT
	ITFSTATESERVER : L_UBUP.L_UBUP_IStateServer;
	ISTATE : INT;
	ECASE : L_UBUP.L_UBUP_StateHandleCase;
END_VAR
END_METHOD

METHOD CHECKTRANSITION
VAR_INPUT
	ITFSTATESERVER : L_UBUP.L_UBUP_IStateServer;
END_VAR
END_METHOD

METHOD DISABLECLIENT : BOOL
VAR_INPUT
	XFIRSTCALL : BOOL;
END_VAR
END_METHOD

METHOD ENABLECLIENT : BOOL
VAR_INPUT
	XFIRSTCALL : BOOL;
END_VAR
END_METHOD

METHOD FINALIZECYCLE
END_METHOD

METHOD LEAVESTATE
END_METHOD

METHOD PREPARECYCLE
END_METHOD

METHOD PREPARESTATECHANGE
END_METHOD

METHOD STIMULATETRANSITION
VAR_INPUT
	ECASE : L_UBUP.L_UBUP_StateHandleCase;
END_VAR
END_METHOD

METHOD UPDATECONDITIONERROR : BOOL
VAR_INPUT
	ITFREQUEST : L_UBUP_IRequest;
END_VAR
END_METHOD

METHOD REQUESTINTERFACE : BOOL
VAR_INPUT
	ID : DINT;
	PITFUNKNOWN : POINTER TO L_UBUP_IUnknown;
END_VAR
END_METHOD

METHOD FB_INIT : BOOL
VAR_INPUT
	BINITRETAINS : BOOL;
	BINCOPYCODE : BOOL;
END_VAR
END_METHOD

METHOD FB_REINIT : BOOL
END_METHOD

METHOD CALL_ALLOCPOINTADR
END_METHOD

METHOD STATE_STANDBY
VAR_INPUT
	ECASE : L_UBUP_StateHandleCase;
	ISTATESERVER : L_UBUP_IStateServer;
END_VAR
END_METHOD

(* ---- L_TB2M_TECHMODULETEMPLATE.pou ---- *)
FUNCTION_BLOCK L_TB2M_TECHMODULETEMPLATE
VAR_INPUT
	XENABLE : BOOL;
	XENABLEOPERATION : BOOL;
	XRESETERROR : BOOL;
	XQSPAPPLICATION : BOOL;
	XABORT : BOOL;
	XJOGPOS : BOOL;
	XJOGNEG : BOOL;
	XHOMEEXECUTE : BOOL;
	LROVERRIDE : LREAL := 1;
	SCCTRLBASICMOTION : L_TB2P_scCtrlBasicMotion;
	SCPAR : L_TB2P_scPar_BasicMotionBase;
END_VAR
VAR_OUTPUT
	XREADYFOROPERATION : BOOL;
	XOPERATIONENABLED : BOOL;
	XREADYFORMOTION : BOOL;
	XERROR : BOOL;
	XWARNING : BOOL;
	EERRORID : L_IE1P_Error;
	XSTOACTIVE : BOOL;
	XQSPACTIVE : BOOL;
	XABORTBUSY : BOOL;
	XABORTDONE : BOOL;
	XJOGGINGBUSY : BOOL;
	XHOMINGBUSY : BOOL;
	XHOMINGDONE : BOOL;
	XISHOMED : BOOL;
	ETMSTATE : L_TB2P_States := L_TB2P_States.DISABLED;
	SCSTATUSBASICMOTION : L_TB2P_scStatusBasicMotion;
	LRSETACCOUT : LREAL;
	LRACTVEL : LREAL;
	LRSETVELOUT : LREAL;
	LRACTPOS : LREAL;
	LRSETPOSOUT : LREAL;
	LRACTFOLLOWINGERROR : LREAL;
END_VAR
VAR_IN_OUT
	AXIS : AXIS_REF;
END_VAR
VAR
	TM_INT : L_TB2M_BasicMotionBase;
	ITFTMSTATECLIENT : L_UBUP_IStateClient;
	ITFSTATESERVER : L_UBUP_IStateServer;
	FB_TRANSITION2STANDBY : L_UBUP_RequestTransitionEdge;
	STATESERVER : L_UBUP_IStateServer;
END_VAR
END_FUNCTION_BLOCK

METHOD EXTENDEDCALLFBS
VAR_INPUT
	ECASE : L_UBUP.L_UBUP_StateHandleCase;
END_VAR
END_METHOD

METHOD EXTENDEDCALLSTATE
VAR_INPUT
	ITFBASE : L_UBUP.L_UBUP_IStateClient;
	ITFSTATESERVER : L_UBUP.L_UBUP_IStateServer;
	ISTATE : INT;
	ECASE : L_UBUP.L_UBUP_StateHandleCase;
END_VAR
END_METHOD

METHOD EXTENDEDCHECKTRANSITION
VAR_INPUT
	ITFSTATESERVER : L_UBUP.L_UBUP_IStateServer;
END_VAR
END_METHOD

METHOD EXTENDEDDISABLECLIENT : BOOL
VAR_INPUT
	XFIRSTCALL : BOOL;
END_VAR
END_METHOD

METHOD EXTENDEDENABLECLIENT : BOOL
VAR_INPUT
	XFIRSTCALL : BOOL;
END_VAR
END_METHOD

METHOD EXTENDEDFINALIZECYCLE
END_METHOD

METHOD EXTENDEDPREPARECYCLE
END_METHOD

METHOD EXTENDEDPREPARESTATECHANGE
END_METHOD

METHOD EXTENDEDSTIMULATETRANSITION
VAR_INPUT
	ECASE : L_UBUP.L_UBUP_StateHandleCase;
END_VAR
END_METHOD

METHOD SETERROR
VAR_INPUT
	XERROR : BOOL;
	EERRORID : L_IE1P_Error;
END_VAR
END_METHOD

METHOD FB_INIT : BOOL
VAR_INPUT
	BINITRETAINS : BOOL;
	BINCOPYCODE : BOOL;
END_VAR
END_METHOD

METHOD LEAVESTATE
END_METHOD

(* ---- L_TB2M_TM_BASE.pou ---- *)
FUNCTION_BLOCK L_TB2M_TM_BASE
VAR_IN_OUT
	INPUT : L_TB2P_BaseIn;
	OUTPUT : L_TB2P_BaseOut;
END_VAR
VAR
	FB_CLIENTPROXY : L_UBUP_StateClientProxy;
	FB_STATESERVER : L_UBUP_StateServer := STRUCT(iFreezeRequestPrio := 10, itfAlternativeRequestByFailedCondition := THIS^);
	ETMSTATE_INT : L_TB2P_States := L_TB2P_States.DISABLED;
	FB_TRANSITION2DISABLED : L_UBUP_RequestTransitionLevel;
	FB_TRANSITION2ERROR : L_UBUP_RequestTransitionLevel;
	FB_TRANSITION2STANDBY : L_UBUP_RequestTransitionEdge;
	ITFSTRUCTPROVIDER : L_TB2P_IStructProvider;
	ITFMCCALLINFOFASSADE : L_UM1P_IMCCallInfo;
	_ITASKIDX : INT;
	_ICALLTASKINDEX : INT;
	_XMULTICOREACTIVE : BOOL;
	_ESUBCOMPTYPE : UDINT;
	_SLICINFO : STRING(10);
	EXTMODULEHANDLER : L_IMHP_IModuleHandler;
	CHILDMODULEHANDLERINT : L_IMHP_IModuleHandler;
	FB_ERRORMANAGER : L_TB2M_ErrorManager;
	ITFERRORMANAGER : L_TB2M_IErrorManager := fb_ErrorManager;
	DWVERSION : DWORD;
	BYCOUNTER : BYTE;
	XHARDWARECHECKPASSED : BOOL;
	XSYSTEMFAULT : BOOL;
	UDIAPPCREDIT : UDINT;
	ICNTRESETERROR : INT := 9;
	XINITDONE : BOOL;
	XEXITDONE : BOOL;
	DIFRAME : DINT;
	DIFRAMESIGNALFLOW : DINT;
	_ITFLENZEVENDORIDCHECKER : L_UBUP_IChecker;
	DECORATOR : L_UBUP_IStateClientDecorator;
	EXTENDEDTECHNOLOGIE : L_UBUP_IStateClientDecorator;
	MONITORSTATESERVER : L_UBUP_IMonitorStateServer;
	STATESERVER : L_UBUP_IStateServer;
END_VAR
END_FUNCTION_BLOCK

METHOD CONNECTCHILD : BOOL
VAR_INPUT
	CHILDMODULEHANDLE : L_IMHP_IModuleHandler;
END_VAR
END_METHOD

METHOD MODULEACTIVATED : BOOL
END_METHOD

METHOD SETADDMODULEINFO
VAR_INPUT
	ESUBCOMPTYPE : UDINT;
	SLICINFO : STRING(10);
END_VAR
END_METHOD

METHOD ERRORSTATUSINFO
VAR_INPUT
	XERROR : BOOL;
	XWARNING : BOOL;
	EERRORID : L_IE1P_Error;
END_VAR
END_METHOD

METHOD HANDOVERRESOURCE : BOOL
VAR_INPUT
	ITFRESOURCE : L_UBUP_IUnknown;
END_VAR
END_METHOD

METHOD ALLOCPOINTADR
VAR_OUTPUT
	IERRORID : INT;
END_VAR
END_METHOD

METHOD HANDLEREJECTEDREQUEST : BOOL
VAR_INPUT
	ITFREQUESTANNOUNCED : L_UBUP_IRequest;
END_VAR
VAR_OUTPUT
	ITFALTERNATIVEREQUEST : L_UBUP_IRequest;
END_VAR
END_METHOD

METHOD CALLFBS
VAR_INPUT
	ECASE : L_UBUP_StateHandleCase;
END_VAR
END_METHOD

METHOD CALLSTATE
VAR_INPUT
	ITFSTATESERVER : L_UBUP_IStateServer;
	ISTATE : INT;
	ECASE : L_UBUP_StateHandleCase;
END_VAR
END_METHOD

METHOD CHECKTRANSITION
VAR_INPUT
	ITFSTATESERVER : L_UBUP_IStateServer;
END_VAR
END_METHOD

METHOD DISABLECLIENT : BOOL
VAR_INPUT
	XFIRSTCALL : BOOL;
END_VAR
END_METHOD

METHOD ENABLECLIENT : BOOL
VAR_INPUT
	XFIRSTCALL : BOOL;
END_VAR
END_METHOD

METHOD FINALIZECYCLE
END_METHOD

METHOD LEAVESTATE
END_METHOD

METHOD PREPARECYCLE
END_METHOD

METHOD PREPARESTATECHANGE
END_METHOD

METHOD STIMULATETRANSITION
VAR_INPUT
	ECASE : L_UBUP_StateHandleCase;
END_VAR
END_METHOD

METHOD UPDATECONDITIONERROR : BOOL
VAR_INPUT
	ITFREQUEST : L_UBUP_IRequest;
END_VAR
END_METHOD

METHOD REQUESTINTERFACE : BOOL
VAR_INPUT
	ID : DINT;
	PITFUNKNOWN : POINTER TO L_UBUP_IUnknown;
END_VAR
END_METHOD

METHOD CALL_CYCLIC
END_METHOD

METHOD STATE_ERROR
VAR_INPUT
	ECASE : L_UBUP_StateHandleCase;
	ITFSTATESERVER : L_UBUP_IStateServer;
END_VAR
END_METHOD

METHOD STATE_EXIT : BOOL
VAR_INPUT
	ECASE : L_UBUP_StateHandleCase;
END_VAR
END_METHOD

METHOD STATE_INIT
VAR_INPUT
	ECASE : L_UBUP_StateHandleCase;
END_VAR
END_METHOD

METHOD STATE_STANDBY
VAR_INPUT
	ECASE : L_UBUP_StateHandleCase;
	ITFSTATESERVER : L_UBUP_IStateServer;
END_VAR
END_METHOD

METHOD FB_REINIT : BOOL
END_METHOD

METHOD FB_INIT : BOOL
VAR_INPUT
	BINITRETAINS : BOOL;
	BINCOPYCODE : BOOL;
	ITFMODULEHANDLER : L_IMHP_IModuleHandler;
END_VAR
END_METHOD

METHOD CALL_HWCHECK : BOOL
END_METHOD

METHOD CALL_SYSTEMFAULT : BOOL
END_METHOD

METHOD CALL_ALLOCPOINTADR
END_METHOD

METHOD CALL_EXIT_CALLFBS
END_METHOD

METHOD CALL_INIT_CALLFBS
END_METHOD

METHOD CALL_RESETOUTPUT
END_METHOD

METHOD MAPTMSTATE
VAR_INPUT
	ETMSTATEINTERNAL : L_TB2P_States;
END_VAR
VAR_OUTPUT
	ETMSTATEEXTERNAL : L_TB2P_States;
END_VAR
END_METHOD

METHOD SETERROR
VAR_INPUT
	XERROR : BOOL;
	EERRORID : L_IE1P_Error;
END_VAR
END_METHOD

(* ---- L_TB2M_TM_MOTIONCONTROL.pou ---- *)
FUNCTION_BLOCK L_TB2M_TM_MOTIONCONTROL EXTENDS L_TB2M_TM_Base
VAR_IN_OUT
	AXIS : AXIS_REF;
END_VAR
VAR
	TM_MOTIONCONTROLCONFIG : L_TB2P_ModuleHandlerConfig;
	XQSPACTIVE_INT : BOOL;
	FB_CONDITIONSTO : L_UBUP_ConditionInput;
	FB_CONDITIONOPERATIONENABLED : L_TB2P_ConditionOperationEnabled;
	FB_CONDITIONLIMITER : L_TB2P_ConditionLimiter;
	FB_CONDITIONAXISNOTSTOPPING : L_TB2P_ConditionAxisNotStopping;
	FB_CONDITIONJOGGINGALLOWEDDIRECTION : L_TB2P_ConditionJogging;
	FB_CONDITIONAXISSTANDSTILL : L_TB2P_ConditionStandstill;
	FB_CONDITIONAXISHOMED : L_UBUP_ConditionInput;
	FB_CONDCOLLECTOPERATIONENABLEDLIMITER : L_UBUP_ConditionCollection := STRUCT(aitfCondition := [fb_ConditionSTO, fb_ConditionOperationEnabled, fb_ConditionLimiter, fb_ConditionAxisNotStopping]);
	FB_CONDCOLLECTOPERATIONENABLEDLIMITERHOMED : L_UBUP_ConditionCollection := STRUCT(aitfCondition := [fb_CondCollectOperationEnabledLimiter, fb_ConditionAxisHomed, fb_ConditionAxisNotStopping]);
	FB_CONDCOLLECTJOGGING : L_UBUP_ConditionCollection := STRUCT(aitfCondition := [fb_ConditionSTO, fb_ConditionOperationEnabled, fb_ConditionLimiter, fb_ConditionJoggingAllowedDirection, fb_ConditionAxisNotStopping]);
	FB_CONDCOLLECTHOMING : L_UBUP_ConditionCollection := STRUCT(aitfCondition := [fb_ConditionSTO, fb_ConditionOperationEnabled, fb_ConditionLimiter, fb_ConditionAxisStandstill]);
	XFORCEABORT : BOOL;
	FB_TRANSITION2QSPAPPL : L_UBUP_RequestTransitionLevel;
	FB_TRANSITION2EXTERNALBYAXIS : L_UBUP_RequestTransitionLevel;
	FB_TRANSITION2STANDYBYAXISDISABLED : L_UBUP_RequestTransitionEdge;
	FB_TRANSITION2HALT : L_UBUP_RequestTransitionEdge;
	FB_TRANSITION2ABORT : L_UBUP_RequestTransitionEdge;
	FB_TRANSITION2EXTERNAL : L_UBUP_RequestTransitionEdge;
	FB_TRANSITION2JOGGING : L_UBUP_RequestTransitionLevel;
	FB_TRANSITION2HOMING : L_UBUP_RequestTransitionEdgeCheckCondition;
	FB_TRANSITION2MOVEVEL : L_UBUP_RequestTransitionEdge;
	FB_TRANSITION2MOVEABS : L_UBUP_RequestTransitionEdge;
	FB_TRANSITION2MOVEREL : L_UBUP_RequestTransitionEdge;
	FB_TRANSITION2MOVEFINISHPOSITIONING : L_UBUP_RequestTransitionEdge;
	PPARMOTIONCTRL : POINTER TO L_TB2P_scPar_TM_MotionControl;
	PSFMOTIONCTRL : POINTER TO L_TB2P_scSF_TM_MotionControl;
	PINPUTBASE : POINTER TO L_TB2P_BasicMotionBaseIn;
	POUTPUTBASE : POINTER TO L_TB2P_BasicMotionBaseOut;
	XSETHOMEPOSSTATEINDEPENDENTACTIVE : BOOL;
	XHOMETRANSITIONNOTBLOCKED : BOOL;
	XHOMEEXECUTE_OLD : BOOL;
	XINTERRUPTHOMINGBYHALT : BOOL;
	FBTEMPLATEABC : L_MC1P_Template;
	PFBTEMPLATEABC : POINTER TO L_MC1P_Template_ForAxis;
	RABC : REFERENCE TO L_MC1P_AxisBasicControl_Internal;
	PAXISINST : POINTER TO AXIS_REF;
	SCDATAABC : L_MC1P_AxisBasicControlInstanceData;
	_XABORTINTERNALNEXTCYLCE : BOOL;
	SCABCIN : L_MC1P_AxisBasicControlInput_Internal;
	SCABCOUT : L_MC1P_AxisBasicControlOutput_Internal;
	XSETJERKDEC : BOOL;
	XJOGGINGSETJERKDEC : BOOL;
	HWLIMITSWITCHINTERFACE : L_MC1P_HWLimitSwitchInterface;
	FB_READAXISINFO : MC_ReadAxisInfo;
	XLIMITERCONTROLVALID : BOOL;
	DWLIMITERCONTROL : DWORD;
	SCDATABASICMOTION : L_TB2P_scDataBasicMotionBase;
	ITFBASICMOTIONBASE : L_TB2P_IBasicMotionBase := THIS^;
	_XUSEBASICMOTIONBASEEXTENSION : BOOL;
	FBHOMINGSTATUS : L_TB2P_BusyDoneManager;
	BASICMOTIONBASEEXTENSION : L_TB2P_IBasicMotionBase;
	CONNECTOR : __SYSTEM.IQueryInterface;
	LRJERKDEC : LREAL;
	LRJOGGINGJERKDEC : LREAL;
	REMAININGTIMEOFPROFILE : LREAL;
	REMAININGTIMEOFPROFILEAVAILABLE : BOOL;
END_VAR
END_FUNCTION_BLOCK

METHOD ALLOCPOINTADR
VAR_OUTPUT
	IERRORID : INT;
END_VAR
END_METHOD

METHOD HANDLEREJECTEDREQUEST : BOOL
VAR_INPUT
	ITFREQUESTANNOUNCED : L_UBUP_IRequest;
END_VAR
VAR_OUTPUT
	ITFALTERNATIVEREQUEST : L_UBUP_IRequest;
END_VAR
END_METHOD

METHOD CALLFBS
VAR_INPUT
	ECASE : L_UBUP_StateHandleCase;
END_VAR
END_METHOD

METHOD CALLSTATE
VAR_INPUT
	ITFSTATESERVER : L_UBUP_IStateServer;
	ISTATE : INT;
	ECASE : L_UBUP_StateHandleCase;
END_VAR
END_METHOD

METHOD CHECKTRANSITION
VAR_INPUT
	ITFSTATESERVER : L_UBUP_IStateServer;
END_VAR
END_METHOD

METHOD FINALIZECYCLE
END_METHOD

METHOD LEAVESTATE
END_METHOD

METHOD PREPARECYCLE
END_METHOD

METHOD STIMULATETRANSITION
VAR_INPUT
	ECASE : L_UBUP_StateHandleCase;
END_VAR
END_METHOD

METHOD STATE_ABORT
VAR_INPUT
	ECASE : L_UBUP_StateHandleCase;
	ITFSTATESERVER : L_UBUP_IStateServer;
END_VAR
END_METHOD

METHOD STATE_EXIT : BOOL
VAR_INPUT
	ECASE : L_UBUP_StateHandleCase;
END_VAR
END_METHOD

METHOD STATE_EXTERNAL
VAR_INPUT
	ECASE : L_UBUP_StateHandleCase;
	ITFSTATESERVER : L_UBUP_IStateServer;
END_VAR
END_METHOD

METHOD STATE_FINISHPOSITIONING
VAR_INPUT
	ECASE : L_UBUP_StateHandleCase;
	ITFSTATESERVER : L_UBUP_IStateServer;
END_VAR
END_METHOD

METHOD STATE_HALT
VAR_INPUT
	ECASE : L_UBUP_StateHandleCase;
	ITFSTATESERVER : L_UBUP_IStateServer;
END_VAR
END_METHOD

METHOD STATE_HOMING
VAR_INPUT
	ECASE : L_UBUP_StateHandleCase;
	ITFSTATESERVER : L_UBUP_IStateServer;
END_VAR
END_METHOD

METHOD STATE_INIT
VAR_INPUT
	ECASE : L_UBUP_StateHandleCase;
END_VAR
END_METHOD

METHOD STATE_JOGGING
VAR_INPUT
	ECASE : L_UBUP_StateHandleCase;
	ITFSTATESERVER : L_UBUP_IStateServer;
END_VAR
END_METHOD

METHOD STATE_MOVEABS
VAR_INPUT
	ECASE : L_UBUP_StateHandleCase;
	ITFSTATESERVER : L_UBUP_IStateServer;
END_VAR
END_METHOD

METHOD STATE_MOVEREL
VAR_INPUT
	ECASE : L_UBUP_StateHandleCase;
	ITFSTATESERVER : L_UBUP_IStateServer;
END_VAR
END_METHOD

METHOD STATE_MOVEVEL
VAR_INPUT
	ECASE : L_UBUP_StateHandleCase;
	ITFSTATESERVER : L_UBUP_IStateServer;
END_VAR
END_METHOD

METHOD STATE_QUICKSTOP
VAR_INPUT
	ECASE : L_UBUP_StateHandleCase;
	ITFSTATESERVER : L_UBUP_IStateServer;
END_VAR
END_METHOD

METHOD CALL_ERRORMANAGER
END_METHOD

METHOD CALL_HWLIMITSWITCH
VAR_INPUT
	ITFTECHMODULE : L_TB2P_IBasicMotionBase;
	XENABLE : BOOL;
	XLIMITSWITCHPOS : BOOL;
	XLIMITSWITCHNEG : BOOL;
END_VAR
VAR_OUTPUT
	XBUSY : BOOL;
	XERROR : BOOL;
	EERRORID : L_IE1P_Error;
END_VAR
END_METHOD

METHOD CALL_READAXISINFO
END_METHOD

METHOD ABCRESETABORT
END_METHOD

METHOD ABCRESETFINISHPOSITIONING
END_METHOD

METHOD ABCRESETHALT
END_METHOD

METHOD ABCRESETHOMEEXECUTE
END_METHOD

METHOD ABCRESETMOVEABSEXECUTE
END_METHOD

METHOD ABCRESETMOVERELEXECUTE
END_METHOD

METHOD ABCRESETMOVEVELEXECUTE
END_METHOD

METHOD CALL_ALLOCPOINTADR
END_METHOD

METHOD CALL_EXIT_CALLFBS
END_METHOD

METHOD CALL_INIT_CALLFBS
END_METHOD

METHOD CALL_RESETOUTPUT
END_METHOD

METHOD MAPTMSTATE
VAR_INPUT
	ETMSTATEINTERNAL : L_TB2P_States;
END_VAR
VAR_OUTPUT
	ETMSTATEEXTERNAL : L_TB2P_States;
END_VAR
END_METHOD

METHOD UPDATEABORTDATA
VAR_INPUT
	LRDEC : LREAL;
	LRJERK : LREAL;
END_VAR
END_METHOD

METHOD CALL_ABC
VAR_INPUT
	ITFTECHMODULE : L_TB2P_IBasicMotionBase;
	XQSPAPPLICATION : BOOL;
	XHALT : BOOL;
	XABORT : BOOL;
	XHOMEEXECUTE : BOOL;
	XJOGPOS : BOOL;
	XJOGNEG : BOOL;
	XFINISHPOSITIONING : BOOL;
	XMOVEVELEXECUTE : BOOL;
	XMOVEABSEXECUTE : BOOL;
	XMOVERELEXECUTE : BOOL;
	XENABLEOPERATION : BOOL;
	XRESETERROR : BOOL;
	XENABLEPOSITIVE : BOOL;
	XENABLENEGATIVE : BOOL;
	XDISABLESWLIMIT : BOOL;
	LROVERRIDE : LREAL;
	LROVERRIDEACC : LREAL;
	LROVERRIDEJERK : LREAL;
	XRESETHOMEPOSITION : BOOL;
	XCONTINUOUSUPDATE : BOOL;
	LRPOS_DIST : LREAL;
	LRVEL : LREAL;
	LRACC : LREAL;
	LRDEC : LREAL;
	LRJERK : LREAL;
	EDIRECTION : MC_DIRECTION;
	SCHOMEEXTTP : MC_TRIGGER_REF;
	XHOMEABSSWITCH : BOOL;
	XSPECIALABORTBEHAVIOR : BOOL;
	LRABORTDEC : LREAL;
	LRABORTJERK : LREAL;
END_VAR
VAR_OUTPUT
	XERROR : BOOL;
	EERRORID : L_IE1P_Error;
	XFUNBUSY : BOOL;
	XFUNDONE : BOOL;
	XFUNCOMMANDABORTED : BOOL;
	EFUNSTATEACT : L_MC1P_ABC_State;
	ECONTROLMODE : L_MC1P_ControlMode;
	XISHOMED : BOOL;
	XHWLIMITSWITCHNEG : BOOL;
	XHWLIMITSWITCHPOS : BOOL;
	XSWLIMITENABLED : BOOL;
	XSWLIMITSWITCHNEG : BOOL;
	XSWLIMITSWITCHPOS : BOOL;
	EAXISTYPE : L_MC1P_DriveType;
	EAXISSTATE : L_MC1P_AXIS_STATE;
	XSTOACTIVE : BOOL;
	XREADYFOROPERATION : BOOL;
	XOPERATIONENABLED : BOOL;
	XREADYFORMOTION : BOOL;
	XAXISWARNING : BOOL;
	XAXISERROR : BOOL;
	EAXISERRORID : L_IE1P_Error;
	XDRIVEWARNING : BOOL;
	XDRIVEERROR : BOOL;
	DWDRIVEERRORID : DWORD;
	LRACTPOS : LREAL;
	LRACTVEL : LREAL;
	LRSETPOSOUT : LREAL;
	LRSETVELOUT : LREAL;
	LRACTFOLLOWINGERROR : LREAL;
	XINPOSITION : BOOL;
	XSTANDSTILLSETVELOCITY : BOOL;
	XSTANDSTILLACTVELOCITY : BOOL;
	XCONSTANTVELOCITY : BOOL;
	XACCELERATING : BOOL;
	XDECELERATING : BOOL;
	XDIRECTIONPOSITIVE : BOOL;
	XDIRECTIONNEGATIVE : BOOL;
	XAXISAVAILABLE : BOOL;
END_VAR
VAR_IN_OUT
	AXIS : AXIS_REF;
END_VAR
END_METHOD

(* ---- L_TB2P_AXISINTERFACE.pou ---- *)
FUNCTION_BLOCK L_TB2P_AXISINTERFACE
VAR_INPUT
	XENABLELIMITSWITCHES : BOOL;
	XENABLEABSHOMESWITCH : BOOL;
	XRELEASEBRAKE : BOOL;
	XSUSPENDANDRESETFOLLOWERROR : BOOL;
	XENABLERESETFOLLOWERROR : BOOL;
	XLOADSPEEDCTRLINTEGRATOR : BOOL;
	LRSPEEDCTRLINTEGRATOR : LREAL := 0;
	XENABLESPEEDPADAPT : BOOL := TRUE;
	LRSPEEDPADAPT : LREAL := 1;
	XENABLEPOSPADAPT : BOOL;
	LRPOSPADAPT : LREAL := 1;
	XENABLEINERTIAADAPT : BOOL;
	LRINERTIAADAPT : LREAL := 1;
	XENABLETORQUEOFFSET : BOOL := FALSE;
	LRTORQUEADD : LREAL := 0;
	XENABLETORQUELIMIT : BOOL := TRUE;
	XACTIVATETORQUELIMITPOS : BOOL;
	XACTIVATETORQUELIMITNEG : BOOL;
	LRTORQUELIMITPOS : LREAL := 2;
	LRTORQUELIMITNEG : LREAL := 2;
	XMONITORINGACTMOTORCURRENT : BOOL := TRUE;
	XMONITORINGDCBUSVOLTAGE : BOOL := TRUE;
	XMONITORINGTHERMALLOADDEVICE : BOOL := TRUE;
	XMONITORINGTHERMALLOADMOTOR : BOOL := TRUE;
	XMONITORINGACTMOTORTEMPERATURE : BOOL := TRUE;
	XMONITORINGSETTORQUE : BOOL := TRUE;
END_VAR
VAR_OUTPUT
	XERROR : BOOL;
	EERRORID : L_IE1P_Error;
	XREADYFORMOTION : BOOL;
	XIMPACTIVE : BOOL;
	XMOTORMAGNETISED : BOOL;
	XVOLTAGEENABLED : BOOL;
	XBRAKERELEASEOUT : BOOL;
	XBRAKERELEASED : BOOL;
	XTORQUELIMITSACTIVE : BOOL;
	XSUSPENDFOLLOWERRORACTIVE : BOOL;
	LRACTTORQUE : LREAL;
	LRACTUALMOTORCURRENT : LREAL;
	LRDC_BUSVOLTAGE : LREAL;
	LRTHERMALLOADDEVICE : LREAL;
	LRTHERMALLOADMOTOR : LREAL;
	LRACTUALMOTORTEMPERATURE : LREAL;
	EAXISSTATE : L_MC1P_Axis_State;
	XLIMITATIONACTIVE : BOOL;
	XLIMITATIONSETTORQUE : BOOL;
	LRACTTORQUESCALED : LREAL;
	XCIA402MODESACTIVE : BOOL;
	LR_ACTSPEED_RPM : LREAL;
	LRSETTORQUE : LREAL;
	WLENZESTATE : WORD;
	WLENZESTATE2 : WORD;
END_VAR
VAR_IN_OUT
	AXIS : AXIS_REF;
END_VAR
VAR
	FB_L_MC1P_BRAKEINTERFACE : L_MC1P_BrakeInterface;
	FB_L_MC1P_SETTORQUELIMIT : L_MC1P_SetTorqueLimit;
	FB_L_MC1P_SETTORQUEOFFSET : L_MC1P_SetTorqueOffset;
	FB_L_MC1P_SUSPENDFOLLOWINGERROR : L_MC1P_SuspendFollowingError;
	FB_L_MC1P_RESETFOLLOWINGERROR : L_MC1P_ResetFollowingError;
	FB_F_TRIG : F_TRIG;
	FB_L_MC1P_SETSPEEDCTRLLOADVALUE : L_MC1P_SetSpeedCtrlLoadValue;
	FB_L_MC1P_SETPOSCTRLADAPTVALUE : L_MC1P_SetPosCtrlAdaptValue;
	FB_L_MC1P_SETSPEEDCTRLADAPTVALUE : L_MC1P_SetSpeedCtrlAdaptValue;
	FB_L_MC1P_SETINERTIAADAPTVALUE : L_MC1P_SetInertiaAdaptValue;
	FB_READACTUALMOTORCURRENT : L_MC1P_CyclicParameterAccessRead;
	FB_READDC_BUSVOLTAGE : L_MC1P_CyclicParameterAccessRead;
	FB_READTHERMALLOADDEVICE : L_MC1P_CyclicParameterAccessRead;
	FB_READTHERMALLOADMOTOR : L_MC1P_CyclicParameterAccessRead;
	FB_READACTUALMOTORTEMPERATURE : L_MC1P_CyclicParameterAccessRead;
	FB_PARREAD_SETTORQUE_0X2DD6_1 : L_MC1P_CyclicParameterAccessRead;
	PAXIS : POINTER TO _AXIS_REF_REAL;
	LRSETTORQUE_SCALED : LREAL;
	LRRATEDTORQUEAXIS : LREAL;
	XINIT : BOOL := TRUE;
END_VAR
END_FUNCTION_BLOCK

METHOD CALL_ERRORHANDLER
END_METHOD

METHOD CALL_FBS
END_METHOD

(* ---- L_TB2P_AXISMOVING.pou ---- *)
FUNCTION_BLOCK L_TB2P_AXISMOVING EXTENDS L_UBUP_ConditionBase
VAR_IN_OUT
	AXIS : AXIS_REF;
END_VAR
END_FUNCTION_BLOCK

METHOD VERIFY : BOOL
VAR_OUTPUT
	XCONDITIONERROR : BOOL;
	EERRORIDPROPOSED : L_IE1P.L_IE1P_Error;
END_VAR
END_METHOD

(* ---- L_TB2P_BASICMOTIONBASE.pou ---- *)
FUNCTION_BLOCK L_TB2P_BASICMOTIONBASE EXTENDS L_TB2P_TechModuleBase
VAR_INPUT
	XENABLE : BOOL;
	XENABLEOPERATION : BOOL;
	XRESETERROR : BOOL;
	XQSPAPPLICATION : BOOL;
	XABORT : BOOL;
	XJOGPOS : BOOL;
	XJOGNEG : BOOL;
	XHOMEEXECUTE : BOOL;
	LROVERRIDE : LREAL := 1;
	SCCTRLBASICMOTION : L_TB2P_scCtrlBasicMotion;
	SCPAR : L_TB2P_scPar_BasicMotionBase;
	SCACCESSPOINTS : L_TB2P_scAP_BasicMotionBase;
END_VAR
VAR_OUTPUT
	XREADYFOROPERATION : BOOL;
	XOPERATIONENABLED : BOOL;
	XREADYFORMOTION : BOOL;
	XERROR : BOOL;
	XWARNING : BOOL;
	EERRORID : L_IE1P_Error;
	XSTOACTIVE : BOOL;
	XQSPACTIVE : BOOL;
	XABORTBUSY : BOOL;
	XABORTDONE : BOOL;
	XJOGGINGBUSY : BOOL;
	XHOMINGBUSY : BOOL;
	XHOMINGDONE : BOOL;
	XISHOMED : BOOL;
	ETMSTATE : L_TB2P_States := L_TB2P_States.DISABLED;
	SCSTATUSBASICMOTION : L_TB2P_scStatusBasicMotion;
	LRACTVEL : LREAL;
	LRSETVELOUT : LREAL;
	LRACTPOS : LREAL;
	LRSETPOSOUT : LREAL;
	LRACTFOLLOWINGERROR : LREAL;
	SCSIGNALFLOW : L_TB2P_scSF_BasicMotionBase;
END_VAR
VAR_IN_OUT
	AXIS : AXIS_REF;
END_VAR
VAR
	TM_INT : L_TB2P_TM_MotionControl := STRUCT(ModuleHandler := ModuleHandler);
	SCPAR_INT : L_TB2P_scPar_BasicMotionBase;
	_UICALLMFUNIDXINPUT : UINT := 1;
	_UICALLMFUNIDXOUTPUT : UINT := 1;
	_ASCINPUT : ARRAY [1.._MCCall.c_BufferDepthInput] OF L_TB2P_BasicMotionBaseIn;
	_ASCOUTPUT : ARRAY [1.._MCCall.c_BufferDepthOutput] OF L_TB2P_BasicMotionBaseOut;
	_ASCPARCORE : ARRAY [1.._MCCall.c_BufferDepthInput] OF L_TB2P_scPar_BasicMotionBase;
	_MCCALL : L_UM1P_MCCall;
	_ASCAP : ARRAY [1.._MCCall.c_BufferDepthInput] OF L_TB2P_scAP_BasicMotionBase;
	_ASCSF : ARRAY [1.._MCCall.c_BufferDepthOutput] OF L_TB2P_scSF_BasicMotionBase;
	_SCACCESSPOINTSCORE : L_TB2P_scAP_BasicMotionBase;
	_SCSIGNALFLOWCORE : L_TB2P_scSF_BasicMotionBase;
	_SCINPUTVISU : L_TB2P_BasicMotionBaseIn;
	_PSCINPUTVISU : POINTER TO L_TB2P_BasicMotionBaseIn := ADR(_scInputVisu);
	_PSCOUTPUTVISU : POINTER TO L_TB2P_BasicMotionBaseOut := ADR(_ascOutput[1]);
	_PSCPARVISU : POINTER TO L_TB2P_scPar_BasicMotionBase := ADR(scPar_int);
	ITFITECHMODULEINTERNAL : L_TB2P_ITechModuleInternal;
	LRJERKDEC : LREAL;
	LRJOGGINGJERKDEC : LREAL;
	REMAININGTIMEOFPROFILE : LREAL;
	REMAININGTIMEOFPROFILEAVAILABLE : BOOL;
END_VAR
END_FUNCTION_BLOCK

METHOD GET_PAP : POINTER TO L_TB2P_scAP_TM_MotionControl
END_METHOD

METHOD GET_PPAR : POINTER TO L_TB2P_scPar_TM_MotionControl
END_METHOD

METHOD GET_PSF : POINTER TO L_TB2P_scSF_TM_MotionControl
END_METHOD

METHOD CALLFUNCTION
VAR_INPUT
	UIINPUTDATAIDX : UINT;
	UIOUTPUTDATAIDX : UINT;
END_VAR
END_METHOD

METHOD COPYINPUTS : BOOL
VAR_INPUT
	IDX : WORD;
END_VAR
END_METHOD

METHOD COPYOUTPUTS : BOOL
VAR_INPUT
	IDX : WORD;
END_VAR
END_METHOD

METHOD FUNCTIONWASCALLEDTWICE : BOOL
VAR_INPUT
	IDX : WORD;
END_VAR
END_METHOD

METHOD HANDLESTANDARDCALL : BOOL
END_METHOD

METHOD SYNCOUTPUTS
VAR_INPUT
	UICOPYOUTPUTFROMIDX : UINT;
	UICOPYOUTPUTTOIDX : UINT;
END_VAR
END_METHOD

METHOD CALL_INTERNALCTRL
END_METHOD

(* ---- L_TB2P_BUSYDONEMANAGER.pou ---- *)
FUNCTION_BLOCK L_TB2P_BUSYDONEMANAGER
VAR
	_XSETBUSY : BOOL;
	_XSETDONE : BOOL;
	_XGETDONE : BOOL;
	_XACKDONE : BOOL;
	BUSY : BOOL;
	DONE : BOOL;
END_VAR
END_FUNCTION_BLOCK

(* ---- L_TB2P_CHECKMODULOOVERRUN.pou ---- *)
FUNCTION_BLOCK L_TB2P_CHECKMODULOOVERRUN
VAR_INPUT
	LRSETPOS : LREAL;
	LRSETVEL : LREAL;
	LRPERIOD : LREAL;
END_VAR
VAR_OUTPUT
	XOVERRUNPOS : BOOL;
	XOVERRUNNEG : BOOL;
END_VAR
VAR
	ALRMEM : ARRAY [1..7] OF LREAL;
	PLRX0 : POINTER TO LREAL;
	PLRX1 : POINTER TO LREAL;
	PLRX2 : POINTER TO LREAL;
	PLRV0 : POINTER TO LREAL;
	PLRV1 : POINTER TO LREAL;
	PLRV2 : POINTER TO LREAL;
	PLRSETVEL_INT : POINTER TO LREAL;
END_VAR
END_FUNCTION_BLOCK

METHOD CALL_CHECKMODULOOVERRUN
VAR_IN_OUT
	LRSETPOS : LREAL;
	LRSETVEL : LREAL;
	LRPERIOD : LREAL;
	XOVERRUNPOS : BOOL;
	XOVERRUNNEG : BOOL;
	ALRMEM : ARRAY [1..7] OF LREAL;
END_VAR
END_METHOD

(* ---- L_TB2P_CLUTCHEXTENDEDBASE.pou ---- *)
FUNCTION_BLOCK L_TB2P_CLUTCHEXTENDEDBASE EXTENDS L_MC2P_ClutchBasic
VAR_INPUT
	XENABLE : BOOL;
	XCLUTCHCLOSE : BOOL;
	XCLUTCHOPENINSTANT : BOOL;
	ECLUTCHMODE : L_TB2P_ClutchMode := L_TB2P_ClutchMode.ramp_pos;
	ECLUTCHDIRECTION : L_MC2P_ClutchDirection := L_MC2P_ClutchDirection.mcCurrentDirection;
	EDIRECTION : L_TB2P_Direction := 0;
	LRCYCMASTERPOS : LREAL;
	LRCYCMASTERVEL : LREAL;
	LRCYCMASTERACC : LREAL;
	LRCYCSLAVEPOS : LREAL;
	LRCYCSLAVEVEL : LREAL;
	LRCYCSLAVEACC : LREAL;
	LROPENINSTANTDEC : LREAL;
	LRMASTERCLOSEPOS : LREAL;
	LRMASTERCLOSEDIST : LREAL := 100;
	LRSLAVECLOSEDIST : LREAL := 100;
	LRMASTEROPENDIST : LREAL := 100;
	LRSLAVEOPENDIST : LREAL := 100;
	LRSLAVEOPENPOS : LREAL;
	LRCLOSETIME : LREAL := 5;
	LROPENTIME : LREAL := 5;
	LRCLUTCHVEL : LREAL := 100;
	LRCLUTCHVELMIN : LREAL := 0;
	LRCLUTCHACC : LREAL := 1000.0;
	LRCLUTCHDEC : LREAL := 1000.0;
	LRCLUTCHJERK : LREAL := 1000000.0;
	LRVELTOLERANCE : LREAL := 1;
	LRAXESCYCLELENGTH : LREAL := 360;
	EMASTERTRAVERSINGRANGE : L_MC1P_TraversingRange;
	LRCYCLETIME : LREAL := 0.001;
	LRSETGROUNDVEL : LREAL := 0;
	LRCYCMASTERVEL_LOCK : LREAL;
END_VAR
VAR_OUTPUT
	XERROR : BOOL;
	EERRORID : L_IE1P_Error;
	XBUSY : BOOL;
	XDONE : BOOL;
	XGROUNDVEL : BOOL;
	XSYNCHRONISED : BOOL;
	XCLUTCHACTIVE : BOOL;
	XWAITOFMASTERTAKESLAVE : BOOL;
	LRSETSLAVEPOSOUT : LREAL;
	LRSETSLAVEVELOUT : LREAL;
	LRSETSLAVEACCOUT : LREAL;
	LRSETSLAVEOFFSETOUT : LREAL;
	LRX0 : LREAL;
	LRX1 : LREAL;
	LRY0 : LREAL;
	LRY1 : LREAL;
	LRX0N : LREAL;
	LRX1N : LREAL;
	LRY0N : LREAL;
	LRY1N : LREAL;
	LRX0P : LREAL;
	LRX1P : LREAL;
	LRY0P : LREAL;
	LRY1P : LREAL;
END_VAR
VAR
	EAXESTRAVERSINGRANGE_INT : L_MC1P_TraversingRange;
	ECLUTCHMODE_INT : L_TB2P_ClutchMode;
	ECLUTCHDIRECTION_LOCK : L_MC2P_ClutchDirection;
	LRVELTOLERANCE_INT : LREAL := 1;
	LRSETSLAVEOFFSET_CLUTCHREL : LREAL;
	LRSETSLAVEOFFSET_INT : LREAL;
	LRSETMASTEROFFSET_OVERRUN : LREAL;
	LRCYCLETIME_INT : LREAL;
	XCLUTCHOPENINSTANT_ACTIVE : BOOL;
	LROPENINSTANTDEC_INT : LREAL;
	XCLUTCHBASICENABLE : BOOL;
	LRTEMP : LREAL;
	LRDELTASETENDPOS : LREAL;
	LRDELTASETENDPOS_OLD : LREAL;
	LRDELTASETENDPOS_OLD2 : LREAL;
	XCLUTCHMASTERVELPOSITIVE : BOOL;
	XMASTERREVERSING : BOOL;
	LRAXESCYCLELENGTH_INT : LREAL;
	XCLUTCHBASIC_EXECUTE_OLD : BOOL;
	XCLUTCHCLOSE_OLD : BOOL;
	XCLUTCHOPENINSTANT_OLD : BOOL;
	XBUSY_OLD : BOOL;
	XENABLE_OLD : BOOL;
	LRCYCMASTERPOS_OLD : LREAL;
	LRMASTERVELADD : LREAL;
	LRMASTERVELADDSYNC : LREAL;
	LRSLAVESTARTPOS : LREAL;
	LRMASTERCLOSEPOS_INT : LREAL;
	LRMASTERCLOSEDIST_INT : LREAL;
	XUSESYNCOUT : BOOL;
	LRSLAVECLOSEDIST_INT : LREAL;
	LRSLAVEOPENDIST_INT : LREAL;
	LRSLAVEOPENPOS_INT : LREAL;
	XSYNCMODEIN_INT : BOOL;
	LRCLUTCHTIME : LREAL;
	LRCYCLECLUTCHTIME : LREAL;
	XCLUTCHPOSMODE_INT : BOOL := TRUE;
	LRCLUTCHVEL_INT : LREAL := 100;
	LRCLUTCHVEL_LOCK : LREAL := 100;
	LRCLUTCHACC_INT : LREAL := 1000.0;
	LRCLUTCHDEC_INT : LREAL := 1000.0;
	LRCLUTCHJERK_INT : LREAL := 1000000.0;
	EMASTERDIRECTION_INT : L_MC2P_ClutchDirection;
	IMASTERMOVEMENTTYPE_INT : INT;
	XREVERSEALLOWED_INT : BOOL;
	XPERIODIC_INT : BOOL;
	LRSLAVEJERK : LREAL;
	ESTATE : L_TB2P_FBStates := L_TB2P_FBStates.INIT;
	XSTATEENTRY : BOOL;
	XSETPARAGAIN : BOOL;
	XERROR_LOCK : BOOL;
	EERRORID_LOCK : L_IE1P_Error;
	LRTOLERANCE : LREAL;
	ICYCLECNTAFTEREXECUTE : INT;
	XRESTART_INT : BOOL;
	SCCYCMASTER : L_MC2P_AxisProfile;
	SCCYCSLAVE : L_MC2P_AxisProfile;
	SCSETSLAVEOUT : L_MC2P_AxisProfile;
	SCSETSLAVEOUT_OLD : L_MC2P_AxisProfile;
	PSCSETSLAVEOUT : POINTER TO L_MC2P_AxisProfile;
	EMASTERDIRECTION : L_MC2P_ClutchDirection;
	XERRORSYNCMODEVELACCREQUIRED : BOOL;
	XERRORINVALIDINPUTDATA : BOOL;
	XCLUTCHBASIC_DONE : BOOL;
	XCLUTCHBASIC_WARNINGCANTPREVENTREVERSE : BOOL;
	XCLUTCHBASIC_ERROR : BOOL;
	ECLUTCHBASIC_ERRORIDCLUTCH : L_IE1P_Error;
	XCLUTCHBASIC_BUSY : BOOL;
	XCLUTCHBASIC_CLUTCHACTIVE : BOOL;
	XCLUTCHBASIC_PERIODIC : BOOL;
	XCLUTCHBASIC_REVERSEALLOWED : BOOL;
	ECLUTCHBASIC_MASTERAXISTYPE : L_MC1P_TraversingRange;
	XCLUTCHBASIC_EXECUTE : BOOL;
	FB_CHECKMODULOOVERRUN : L_TB2P_CheckModuloOverrun;
	XHALT_OLD : BOOL;
	XHALTBUSYINT : BOOL;
	XHALTDONEINT : BOOL;
	LRHALTTIME : LREAL;
	LRHALTDIST : LREAL;
	_IDX1 : INT;
	_IDX2 : INT;
	_LRFACTOR : LREAL;
	_LRFACTORINV : LREAL;
	_XADAPTSLAVE : BOOL;
	_LRSLAVEPOS : LREAL;
	XSIMPLEFUNRAMPSLAVEDIST : BOOL := TRUE;
	LRSETSLAVEOFFSET_CLUTCHRELENTRY : LREAL;
	SCCYCSLAVE_CLUTCHRELENTRY : L_MC2P_AxisProfile;
	XRAMPDISTABSVIALINEAR : BOOL;
	XCLUTCHBASIC_BUSY_OLD : BOOL;
	XCLUTCHMASTERVELPOSITIVE_OLD : BOOL;
	XMASTERINSIDEXSIZE : BOOL;
	XMASTERINSIDEXSIZE_OLD : BOOL;
	XMASTERINSIDEXSIZEP : BOOL;
	XMASTERINSIDEXSIZEP_OLD : BOOL;
	XMASTERINSIDEXSIZEN : BOOL;
	XMASTERINSIDEXSIZEN_OLD : BOOL;
	XCLUTCHDIRECTIONPOSITIVE : BOOL;
	ALRKOEF : ARRAY [0..5] OF LREAL;
	LRXFACTORN : LREAL;
	LRYFACTORN : LREAL;
	LRSETSLAVEOFFSET_CLUTCHRELN : LREAL;
	LRXFACTORP : LREAL;
	LRYFACTORP : LREAL;
	LRSETSLAVEOFFSET_CLUTCHRELP : LREAL;
	LRXFACTOR : LREAL;
	LRYFACTOR : LREAL;
	LRXSCALED : LREAL;
	LRYSCALED : LREAL;
	LRYSCALED_OLD : LREAL;
	LRYSCALEDDIFF : LREAL;
	LRSETYPOS : LREAL;
	LRSETYPOS_OLD : LREAL;
	LRSETYVEL : LREAL;
	LRSETYVEL_OLD : LREAL;
	LRSETYACC : LREAL;
	XCLUTCHDIRECTIONPOSITIVE_OLD : BOOL;
	LRMASTERCYCLELENGTH : LREAL;
	LRDUMMY : LREAL;
	LRCYCMASTERVEL_OLD : LREAL;
	WRAMPVELLACCSTEPPER : WORD;
	XNOREVERSEACTIVE : BOOL;
	XHALT_BUSY : BOOL;
	XHALT_DONE : BOOL;
	XSLAVEHALT : BOOL;
	XSLAVEHALT_OLD : BOOL;
	EALLOWEDDIRECTION_INT : L_TB2P_AllowedDirection;
	XWAITOFMASTERALLOWEDDIRECTION : BOOL;
	XWAITOFMASTERALLOWEDDIRECTION_OLD : BOOL;
	XSYNCHRONISED_OLD : BOOL;
	LRSETGROUNDVEL_LOCK : LREAL := 0;
	LRGROUNDVELDIFFVEL_LOCK : LREAL := 0;
	LRGROUNDVELSTARTVEL_LOCK : LREAL := 0;
	LRSETYPOSADDITIONAL : LREAL;
	SCCYCMASTERATGROUNDVEL : L_MC2P_AxisProfile;
	LRSTARTVELFAKTOR : LREAL;
	LRVELFACTOR : LREAL;
	LRYDISTSCALED : LREAL;
	XSYNCINSTANDSTILLMASTER : BOOL;
	LRWAITMASTERDIST : LREAL;
	XWAITOFMASTER : BOOL;
	XWAITAFTERREACHEDSTANDSTILL : BOOL;
	XSYNCOVERSPEED : BOOL := FALSE;
	XSYNCUNDERSPEED : BOOL := FALSE;
	XSTARTVELATENABLE : BOOL;
	AIMASTERDIRECTION : ARRAY [0..2] OF INT;
	IMASTERDIRECTION : INT;
	ICOUNTER : INT;
	ICOUTERMAX : INT := 15;
	XRESTARTSYNCIN : BOOL;
	LRMASTERVELATEXECUTE : LREAL;
	XSYNCINASFLYINGSAW : BOOL;
	FB_STACKCONTROLARRAYNOISE : L_MC1P_StackControlArray := STRUCT(iMaxLegth := 10);
	ALRDELTAVEL : ARRAY [0..10] OF LREAL;
	AXNOISE : ARRAY [0..5] OF BOOL;
	ALRVELTOLERANCE : ARRAY [0..5] OF LREAL;
	XNOISE : BOOL;
	XACCPOSITIV : BOOL;
	IACCCHANGEDIRECTIONCOUNTER : INT;
	XOPENONLIMIT_INT : BOOL;
	XCLUTCHOLD2 : BOOL;
	C_ALRKOEF_SYNCIN : ARRAY [0..5] OF LREAL := [0, 0, 0, 1, -0.5, 0];
	C_ALRKOEF_SYNCOUT : ARRAY [0..5] OF LREAL := [0, 1, 0, -1, 0.5, 0];
	C_ALRKOEF_0_1 : ARRAY [0..5] OF LREAL := [0, 0, 0, 10, -15, 6];
END_VAR
END_FUNCTION_BLOCK

METHOD CALL_ALLOCPOINTADR
END_METHOD

METHOD CALL_CHECKMASTERNOISE : BOOL
END_METHOD

METHOD CALL_CLUTCHCLOSEMODE
END_METHOD

METHOD CALL_CLUTCHOPENMODE
END_METHOD

METHOD CALL_ERRORHANDLER
END_METHOD

METHOD CALL_FBMETHODS
END_METHOD

METHOD CALL_FB_CHECKMODULOOVERRUN
END_METHOD

METHOD CALL_FB_CLUTCHBASIC_GROUNDVEL_RAMPPOS
END_METHOD

METHOD CALL_FB_CLUTCHBASIC_GROUNDVEL_VELLACC
END_METHOD

METHOD CALL_FB_CLUTCHBASIC_OPENINSTANT
END_METHOD

METHOD CALL_FB_CLUTCHBASIC_RAMPABS
END_METHOD

METHOD CALL_FB_CLUTCHBASIC_RAMPABS_TARGETPOS
END_METHOD

METHOD CALL_FB_CLUTCHBASIC_RAMPPOS
END_METHOD

METHOD CALL_FB_CLUTCHBASIC_RAMPREL
END_METHOD

METHOD CALL_FB_CLUTCHBASIC_RAMPTIME
END_METHOD

METHOD CALL_FB_CLUTCHBASIC_RAMPVELLACC
END_METHOD

METHOD CALL_FB_CLUTCHBASIC_RELATIVE
END_METHOD

METHOD CALL_MASTERDIRECTION
END_METHOD

METHOD CALL_MODULOTOLINEARMASTERPOS
END_METHOD

METHOD CALL_OPENONLIMITED
VAR_IN_OUT
	XCLUTCH : BOOL;
	SCINPUTSLAVE : L_MC2P_AxisProfile;
	XPOSMODE : BOOL;
	LRSLAVEOPENPOS : LREAL;
	LRMAXVELDIFF : LREAL;
	LRMAXACC : LREAL;
	LRMAXDEC : LREAL;
	LRJERK : LREAL;
	LRCYCLETIME : LREAL;
	SCOUTPUTSLAVE : L_MC2P_AxisProfile;
	XBUSY : BOOL;
	XDONE : BOOL;
	XERROR : BOOL;
	EERRORID : L_IE1P_Error;
END_VAR
END_METHOD

METHOD CALL_OUTPUT
END_METHOD

METHOD CALL_RAMPRELDIESTREL_CALCCOEFX0X1Y0Y1
END_METHOD

METHOD CALL_RAMPRELDISTABS_CALCCOEFX0X1Y0Y1
END_METHOD

METHOD CALL_RAMPRELDISTABS_CORRX0X1FORMODULOMASTER
END_METHOD

METHOD CALL_RAMPSLAVEDIST_ABS
END_METHOD

METHOD CALL_RAMPSLAVEDIST_REL
END_METHOD

METHOD CALL_RAMPSLAVEDIST_SETYPOSOUT
END_METHOD

METHOD CALL_RAMPSLAVETIME_SETYPOSOUT
END_METHOD

METHOD CALL_RESETCLUTCH
END_METHOD

METHOD CALL_RESETCOMMANDS
END_METHOD

METHOD CALL_RESETOUTPUT
END_METHOD

METHOD CALL_SETCLUTCHCLOSEPAR
END_METHOD

METHOD CALL_SETCLUTCHCLOSEPAR_VELACC
END_METHOD

METHOD CALL_SETCLUTCHOPENPAR
END_METHOD

METHOD CALL_STATEMASHINE
END_METHOD

METHOD CALL_WAITOFMASTERALLOWEDDIRECTION
END_METHOD

METHOD SET_CLUTCHOFFSET : BOOL
VAR_INPUT
	LRIN : LREAL := 0;
END_VAR
END_METHOD

METHOD SLAVEHALT
VAR_INPUT
	XHALT : BOOL;
	SCACTSLAVE : L_MC2P_AxisProfile;
	LRMAXVELDIFF : LREAL;
	LRMAXACC : LREAL;
	LRMAXDEC : LREAL;
	LRJERK : LREAL;
	LRCYCLETIME : LREAL;
END_VAR
VAR_OUTPUT
	SCOUTPUTSLAVE : L_MC2P_AxisProfile;
	XBUSY : BOOL;
	XDONE : BOOL;
	XERROR : BOOL;
	EERRORID : L_IE1P_Error;
END_VAR
END_METHOD

METHOD CALL_S000_CYCLIC
END_METHOD

METHOD CALL_S001_INIT
END_METHOD

METHOD CALL_S010_READY
END_METHOD

METHOD CALL_S051_GROUNDSPEED
END_METHOD

METHOD CALL_S100_CLUTCH_CLOSE
END_METHOD

METHOD CALL_S200_SYNCHRON
END_METHOD

METHOD CALL_S300_CLUTCH_OPEN
END_METHOD

METHOD CALL_S998_ERROR
END_METHOD

(* ---- L_TB2P_CONDITIONAXISNOTSTOPPING.pou ---- *)
FUNCTION_BLOCK L_TB2P_CONDITIONAXISNOTSTOPPING EXTENDS L_UBUP_ConditionBase
VAR_IN_OUT
	AXIS : AXIS_REF;
END_VAR
END_FUNCTION_BLOCK

METHOD VERIFY : BOOL
VAR_OUTPUT
	XCONDITIONERROR : BOOL;
	EERRORIDPROPOSED : L_IE1P.L_IE1P_Error;
END_VAR
END_METHOD

(* ---- L_TB2P_CONDITIONBASEVELOCITYDIRECTION.pou ---- *)
FUNCTION_BLOCK L_TB2P_CONDITIONBASEVELOCITYDIRECTION EXTENDS L_UBUP_ConditionBase
VAR_INPUT
	LRBASEVELOCITY : LREAL;
	EALLOWEDDIR : L_TB2P_AllowedDirection;
	DWLIMITERCONTROL : DWORD;
END_VAR
VAR_OUTPUT
	XDIRECTIONDISABLED : BOOL;
	XINVALIDINPUT : BOOL;
END_VAR
VAR_IN_OUT
	AXIS : AXIS_REF;
END_VAR
END_FUNCTION_BLOCK

METHOD VERIFY : BOOL
VAR_OUTPUT
	XCONDITIONERROR : BOOL;
	EERRORIDPROPOSED : L_IE1P.L_IE1P_Error;
END_VAR
END_METHOD

(* ---- L_TB2P_CONDITIONGT.pou ---- *)
FUNCTION_BLOCK L_TB2P_CONDITIONGT EXTENDS L_UBUP_ConditionBase
VAR_INPUT
	LRVALUE : LREAL;
	LRTARGET : LREAL;
END_VAR
VAR
	ECONDITIONWARNINGID_INT : L_IE1P_Error;
END_VAR
END_FUNCTION_BLOCK

METHOD VERIFY : BOOL
VAR_OUTPUT
	XCONDITIONERROR : BOOL;
	EERRORIDPROPOSED : L_IE1P.L_IE1P_Error;
END_VAR
END_METHOD

METHOD FB_INIT : BOOL
VAR_INPUT
	BINITRETAINS : BOOL;
	BINCOPYCODE : BOOL;
	ECONDITIONWARNINGID : L_IE1P_Error;
END_VAR
END_METHOD

(* ---- L_TB2P_CONDITIONJOGGING.pou ---- *)
FUNCTION_BLOCK L_TB2P_CONDITIONJOGGING EXTENDS L_UBUP_ConditionBase
VAR_INPUT
	XJOGPOS : BOOL;
	XJOGNEG : BOOL;
	DWLIMITERCONTROL : DWORD;
END_VAR
VAR_OUTPUT
	XDIRECTIONDISABLED : BOOL;
	XINVALIDINPUT : BOOL;
END_VAR
VAR_IN_OUT
	AXIS : AXIS_REF;
END_VAR
END_FUNCTION_BLOCK

METHOD VERIFY : BOOL
VAR_OUTPUT
	XCONDITIONERROR : BOOL;
	EERRORIDPROPOSED : L_IE1P.L_IE1P_Error;
END_VAR
END_METHOD

(* ---- L_TB2P_CONDITIONLIMITER.pou ---- *)
FUNCTION_BLOCK L_TB2P_CONDITIONLIMITER EXTENDS L_UBUP_ConditionBase
VAR_INPUT
	DWLIMITERCONTROL : DWORD;
END_VAR
END_FUNCTION_BLOCK

METHOD VERIFY : BOOL
VAR_OUTPUT
	XCONDITIONERROR : BOOL;
	EERRORIDPROPOSED : L_IE1P.L_IE1P_Error;
END_VAR
END_METHOD

(* ---- L_TB2P_CONDITIONMASTERDIRECTION.pou ---- *)
FUNCTION_BLOCK L_TB2P_CONDITIONMASTERDIRECTION EXTENDS L_UBUP_ConditionBase
VAR_INPUT
	MASTERVALUES : L_MC1P_IAXIS_REF_MASTERVALUES;
	EALLOWEDDIR : L_TB2P_AllowedDirection;
	DWLIMITERCONTROL : DWORD;
END_VAR
VAR_OUTPUT
	XDIRECTIONDISABLED : BOOL;
	XINVALIDINPUT : BOOL;
END_VAR
VAR_IN_OUT
	AXIS : AXIS_REF;
END_VAR
END_FUNCTION_BLOCK

METHOD VERIFY : BOOL
VAR_OUTPUT
	XCONDITIONERROR : BOOL;
	EERRORIDPROPOSED : L_IE1P.L_IE1P_Error;
END_VAR
END_METHOD

(* ---- L_TB2P_CONDITIONOPERATIONDISABLED.pou ---- *)
FUNCTION_BLOCK L_TB2P_CONDITIONOPERATIONDISABLED EXTENDS L_UBUP_ConditionBase
VAR_IN_OUT
	AXIS : AXIS_REF;
END_VAR
END_FUNCTION_BLOCK

METHOD VERIFY : BOOL
VAR_OUTPUT
	XCONDITIONERROR : BOOL;
	EERRORIDPROPOSED : L_IE1P.L_IE1P_Error;
END_VAR
END_METHOD

(* ---- L_TB2P_CONDITIONOPERATIONENABLED.pou ---- *)
FUNCTION_BLOCK L_TB2P_CONDITIONOPERATIONENABLED EXTENDS L_UBUP_ConditionBase
VAR_IN_OUT
	AXIS : AXIS_REF;
END_VAR
END_FUNCTION_BLOCK

METHOD VERIFY : BOOL
VAR_OUTPUT
	XCONDITIONERROR : BOOL;
	EERRORIDPROPOSED : L_IE1P.L_IE1P_Error;
END_VAR
END_METHOD

(* ---- L_TB2P_CONDITIONSTANDSTILL.pou ---- *)
FUNCTION_BLOCK L_TB2P_CONDITIONSTANDSTILL EXTENDS L_UBUP_ConditionBase
VAR_IN_OUT
	AXIS : AXIS_REF;
END_VAR
END_FUNCTION_BLOCK

METHOD VERIFY : BOOL
VAR_OUTPUT
	XCONDITIONERROR : BOOL;
	EERRORIDPROPOSED : L_IE1P.L_IE1P_Error;
END_VAR
END_METHOD

(* ---- L_TB2P_CONDITIONSTATENOTJOGGING.pou ---- *)
FUNCTION_BLOCK L_TB2P_CONDITIONSTATENOTJOGGING EXTENDS L_UBUP_ConditionBase
VAR_IN_OUT
	ETMSTATEINTERNAL : L_TB2P_States;
END_VAR
END_FUNCTION_BLOCK

METHOD VERIFY : BOOL
VAR_OUTPUT
	XCONDITIONERROR : BOOL;
	EERRORIDPROPOSED : L_IE1P.L_IE1P_Error;
END_VAR
END_METHOD

(* ---- L_TB2P_CTRLBASICMOTION.pou ---- *)
FUNCTION_BLOCK L_TB2P_CTRLBASICMOTION
VAR_INPUT
	XENABLEPOSITIVE : BOOL := TRUE;
	XENABLENEGATIVE : BOOL := TRUE;
	LROVERRIDEACC : LREAL := 1;
	LROVERRIDEJERK : LREAL := 1;
	XDISABLESWLIMIT : BOOL;
	XCONTINUOUSUPDATE : BOOL := TRUE;
	XHALT : BOOL;
	XFINISHPOSITIONING : BOOL;
	XMOVEVELEXECUTE : BOOL;
	XMOVEABSEXECUTE : BOOL;
	XMOVERELEXECUTE : BOOL;
	LRPOS_DIST : LREAL := 0;
	XHOMEABSSWITCH : BOOL;
	XRESETHOMEPOSITION : BOOL;
	XHWLIMITPOS : BOOL;
	XHWLIMITNEG : BOOL;
END_VAR
VAR_OUTPUT
	SCCTRLBASICMOTION : L_TB2P_scCtrlBasicMotion;
END_VAR
END_FUNCTION_BLOCK

(* ---- L_TB2P_FBBASENOAXIS.pou ---- *)
FUNCTION_BLOCK L_TB2P_FBBASENOAXIS EXTENDS L_MC1P_Template_NoAxis
END_FUNCTION_BLOCK

(* ---- L_TB2P_GETAXISVALUES_BASE.pou ---- *)
FUNCTION_BLOCK L_TB2P_GETAXISVALUES_BASE
VAR_OUTPUT
	LRAXISCYCLELENGTH : LREAL;
	LRAXISSETPOSITION : LREAL;
	LRAXISSETVELOCITY : LREAL;
	LRAXISSETACCELERATION : LREAL;
	LRAXISSETTORQUE : LREAL;
END_VAR
VAR_IN_OUT
	AXIS : AXIS_REF;
END_VAR
END_FUNCTION_BLOCK

(* ---- L_TB2P_GETMASTERVALUEDIRECTION.pou ---- *)
FUNCTION_BLOCK L_TB2P_GETMASTERVALUEDIRECTION
VAR_INPUT
	LRCYCSETPOSIN : LREAL;
	LRCYCSETVELIN : LREAL;
	ETRAVERSINGRANGE : L_MC1P_TraversingRange;
	LRCYCLELENGTH : LREAL;
END_VAR
VAR_OUTPUT
	XPOSITIVE : BOOL := FALSE;
	XNEGATIVE : BOOL := FALSE;
	XSTANDSTILL : BOOL := TRUE;
END_VAR
VAR
	LRPOSDIFF : LREAL;
	ALRPOSDIFF : ARRAY [1..10] OF LREAL := [0, 0, 0, 0, 0, 0, 0, 0, 0, 0];
	BYCOUNTER : BYTE := 1;
	LRCYCSETPOSIN_OLD : LREAL;
	I : BYTE := 1;
	LRSUMMEPOSDIFF : LREAL;
	XFIRSTCYCLESTANDSTILL : BOOL := TRUE;
	LRPOSITIONSTANDSTILL : LREAL;
	LRTHRESHOLDPOS : LREAL;
	LRTHRESHOLDNEG : LREAL;
	XPOSITIVEDRIFT : BOOL;
	XNEGATIVEDRIFT : BOOL;
	LRMIN : LREAL;
	LRMAX : LREAL;
	LRHYST : LREAL;
	XHYSTFOUND : BOOL;
	LRVARIANCE : LREAL := 1E-06;
	LRTMPMIN : LREAL;
	LRTMPMAX : LREAL;
	ICOUNT : INT;
	XINITDONE : BOOL := FALSE;
	LRMITTELWERT_ENCODER : LREAL;
	XOPERATIONENABLEDOLD : BOOL;
	LRVELDIFF : LREAL;
	LRFACTOR : LREAL := 500;
	LRFACTOR_INT : LREAL;
	XENCODERCHANGE : BOOL := FALSE;
	LRMITTELWERT : LREAL := 0;
	XOPERATIONENABLED : BOOL;
	CLRVARIANCE : LREAL := 1E-09;
END_VAR
END_FUNCTION_BLOCK

METHOD ISBETWEEN : BOOL
VAR_INPUT
	LRVALUE : LREAL;
	LRUPPER : LREAL;
	LRLOWER : LREAL;
	LRVARIANCE : LREAL := 1E-09;
END_VAR
END_METHOD

METHOD ISOUTSIDE : BOOL
VAR_INPUT
	LRVALUE : LREAL;
	LRUPPER : LREAL;
	LRLOWER : LREAL;
	LRVARIANCE : LREAL := 1E-09;
END_VAR
END_METHOD

(* ---- L_TB2P_GETMASTERVALUES_BASE.pou ---- *)
FUNCTION_BLOCK L_TB2P_GETMASTERVALUES_BASE
VAR_INPUT
	AXIS : L_MC1P_IAXIS_REF_MASTERVALUES;
END_VAR
VAR_OUTPUT
	LRAXISCYCLELENGTH : LREAL;
	LRAXISSETPOSITION : LREAL;
	LRAXISSETVELOCITY : LREAL;
	LRAXISSETACCELERATION : LREAL;
	LRAXISSETTORQUE : LREAL;
END_VAR
END_FUNCTION_BLOCK

(* ---- L_TB2P_MODULEHANDLERCONFIG.pou ---- *)
FUNCTION_BLOCK L_TB2P_MODULEHANDLERCONFIG
END_FUNCTION_BLOCK

METHOD FB_INIT : BOOL
VAR_INPUT
	BINITRETAINS : BOOL;
	BINCOPYCODE : BOOL;
	ITFTM_BASE : L_TB2P_ITM_Base;
	ESUBCOMPTYPE : UDINT;
	SLICENSE : STRING(10);
END_VAR
END_METHOD

(* ---- L_TB2P_SETAXISREF.pou ---- *)
FUNCTION_BLOCK L_TB2P_SETAXISREF
VAR_INPUT
	ETRAVERSINGRANGE : L_MC1P_TraversingRange;
	LRAXISCYCLELENGTH : LREAL;
	LRAXISSETPOSITION : LREAL;
	LRAXISSETVELOCITY : LREAL;
	LRAXISSETACCELERATION : LREAL;
	LRAXISSETTORQUE : LREAL;
END_VAR
VAR_OUTPUT
	MASTERAXIS : L_MC1P_IAXIS_REF_MASTERVALUES;
END_VAR
VAR
	MASTERVALUES : L_MC1P_SetAxisRefMasterValues;
	XERRORINVALIDCYCLELENGTH : BOOL;
END_VAR
END_FUNCTION_BLOCK

(* ---- L_TB2P_SETTORQUELIMIT.pou ---- *)
FUNCTION_BLOCK L_TB2P_SETTORQUELIMIT
VAR_INPUT
	ESELECTIONEXTTORQUELIMIT : L_TB2P_eSelectionExtTorqueLimit;
	XENABLEEXTERNALTORQUELIMIT : BOOL;
	LREXTERNALTORQUELIMIT : LREAL;
END_VAR
VAR_OUTPUT
	XENABLETORQUELIMITPOSOUT : BOOL;
	XENABLETORQUELIMITNEGOUT : BOOL;
	LRTORQUELIMITPOSOUT : LREAL;
	LRTORQUELIMITNEGOUT : LREAL;
END_VAR
END_FUNCTION_BLOCK

(* ---- L_TB2P_SOURCEMONITORINGSIGNALS.pou ---- *)
FUNCTION_BLOCK L_TB2P_SOURCEMONITORINGSIGNALS
VAR_INPUT
	LRACTUALMOTORTEMPERATURE : LREAL;
	LRACTUALMOTORCURRENT : LREAL;
	LRDCBUSVOLTAGE : LREAL;
	LRTHERMALLOADDEVICE : LREAL;
	LRTHERMALLOADMOTOR : LREAL;
	IANALOGSIGNAL : INT;
END_VAR
VAR_OUTPUT
	DWMONITORINGSIGNALS : DWORD;
END_VAR
END_FUNCTION_BLOCK

METHOD CALL_SOURCEMONITORINGSIGNALS : DWORD
END_METHOD

(* ---- L_TB2P_STATUSBASICMOTION.pou ---- *)
FUNCTION_BLOCK L_TB2P_STATUSBASICMOTION
VAR_INPUT
	SCSTATUSBASICMOTION : L_TB2P_scStatusBasicMotion;
END_VAR
VAR_OUTPUT
	XFUNBUSY : BOOL;
	XFUNDONE : BOOL;
	XFUNCOMMANDABORTED : BOOL;
	XHALTBUSY : BOOL;
	XHALTDONE : BOOL;
	ECONTROLMODE : L_MC1P_ControlMode;
	XHWLIMITSWITCHNEG : BOOL;
	XHWLIMITSWITCHPOS : BOOL;
	XSWLIMITENABLED : BOOL;
	XSWLIMITSWITCHNEG : BOOL;
	XSWLIMITSWITCHPOS : BOOL;
	EAXISTYPE : L_MC1P_DriveType;
	EAXISSTATE : L_MC1P_AXIS_STATE;
	XAXISWARNING : BOOL;
	XAXISERROR : BOOL;
	XDRIVEWARNING : BOOL;
	XDRIVEERROR : BOOL;
	DWDRIVEERRORID : DWORD;
	XCONSTANTVELOCITY : BOOL;
	XACCELERATING : BOOL;
	XDECELERATING : BOOL;
	XDIRECTIONPOSITIVE : BOOL;
	XDIRECTIONNEGATIVE : BOOL;
	XINPOSITION : BOOL;
	XAXISAVAILABLE : BOOL;
	XSTANDSTILLSETVELOCITY : BOOL;
	XSTANDSTILLACTVELOCITY : BOOL;
END_VAR
END_FUNCTION_BLOCK

(* ---- L_TB2P_SYNCMOTIONCONTROL.pou ---- *)
FUNCTION_BLOCK L_TB2P_SYNCMOTIONCONTROL EXTENDS L_TB2P_TM_MotionControl
VAR_INPUT
	MASTERVALUES : L_MC1P_IAXIS_REF_MASTERVALUES;
END_VAR
VAR
	MASTERVALUES_INT : L_MC1P_IAXIS_REF_MASTERVALUES;
	XMASTERITFVALID : BOOL;
	BYMASTERID : POINTER TO BYTE;
	XMASTERITFVALID_LOCK : BOOL;
	BYMASTERID_LOCK : POINTER TO BYTE;
	XTMNEEDSNOMASTERREF : BOOL;
END_VAR
END_FUNCTION_BLOCK

METHOD CALL_ALLOCPOINTADR
END_METHOD

METHOD CALL_ERRORHANDLER
END_METHOD

METHOD CALL_MASTERAXISREF
VAR_INPUT
	MASTERVALUES : L_MC1P_IAXIS_REF_MASTERVALUES;
END_VAR
END_METHOD

(* ---- L_TB2P_TECHMODULEBASE.pou ---- *)
FUNCTION_BLOCK L_TB2P_TECHMODULEBASE
VAR
	MODULEHANDLERBASE : L_IMHP_ModuleHandler := STRUCT(UseLEM := TRUE, CompActiveDefault := TRUE, Layer := L_IMHP_Layer.Tech_Application, CompType := L_IMHP_ComponentType.TechnologyModule);
	_FBVENDORIDCHECKER : L_UBUP_VendorIdChecker;
	_ITFLENZEVENDORIDCHECKER : L_UBUP_IChecker := _fbVendorIdChecker;
	XINTERNALCONTROL : BOOL;
	XINTERNALCONTROLACTIVE : BOOL;
	DIFRAME : DINT;
	DIFRAMESIGNALFLOW : DINT;
	_ITASKIDX : INT;
	HWCHECKER : L_UBUP_IChecker;
	ITFITECHMODULEINTERNAL : L_TB2P_ITechModuleInternal;
	MODULEHANDLER : L_IMHP_IModuleHandler;
	TASKIDX : INT;
END_VAR
END_FUNCTION_BLOCK

METHOD MODULEDISABLED
END_METHOD

METHOD MODULEENABLED
VAR_INPUT
	CHILDMODULEHANDLE : L_IMHP_IModuleHandler;
END_VAR
END_METHOD

METHOD GET_PAP : POINTER TO L_TB2P_scAP_TM_MotionControl
END_METHOD

METHOD GET_PPAR : POINTER TO L_TB2P_scPar_TM_MotionControl
END_METHOD

METHOD GET_PSF : POINTER TO L_TB2P_scSF_TM_MotionControl
END_METHOD

METHOD REQUESTINTERFACE : BOOL
VAR_INPUT
	ID : DINT;
	PITFUNKNOWN : POINTER TO L_UBUP.L_UBUP_IUnknown;
END_VAR
END_METHOD

METHOD FB_AFTERINIT : BOOL
END_METHOD

(* ---- L_TB2P_TM_BASE.pou ---- *)
FUNCTION_BLOCK L_TB2P_TM_BASE
VAR_INPUT
	CHILDMODULE : L_IMHP_IModuleHandler;
END_VAR
VAR_IN_OUT
	INPUT : L_TB2P_BaseIn;
	OUTPUT : L_TB2P_BaseOut;
END_VAR
VAR
	ITFSTRUCTPROVIDER : L_TB2P_IStructProvider;
	DWVERSION : DWORD;
	DWVENDORID : DWORD;
	BYCOUNTER : BYTE;
	XHARDWARECHECKPASSED : BOOL;
	XSYSTEMFAULT : BOOL;
	UDIAPPCREDIT : UDINT;
	XABCINTERNALCONTROLACTIVE : BOOL;
	XENABLE_OLD : BOOL;
	XENABLE_LOCK : BOOL;
	XRESETERROR_OLD : BOOL := FALSE;
	XRESETERRORINIT : BOOL;
	XTMWARNING_INT : BOOL;
	XTMWARNING_OLD : BOOL;
	XTMERROR_INT : BOOL;
	XTMERROR_OLD : BOOL;
	ETMERRORID_INT : L_IE1P_Error;
	ETMERRORID_OLD : L_IE1P_Error;
	XERROR_FIRST : BOOL;
	EERRORID_FIRST : L_IE1P_Error;
	XRESETERROR_RTRIG : BOOL;
	XRESETOUTPUTDONE : BOOL;
	_IRESETOUTPUTCNTRCYCLES : INT;
	XERROR_OLD : BOOL;
	XWARNING_OLD : BOOL;
	ICNTRESETERROR : INT := 10;
	XINITDONE : BOOL;
	XINITDONE_OLD : BOOL;
	IINITSTATE : INT;
	XTMENABLED : BOOL;
	REQUESTSINFO : DWORD;
	REQUESTSINFO_OLD : DWORD;
	DWRTRIG : DWORD;
	XNEWREQUEST : BOOL;
	XREQUEST_FTRIG : BOOL;
	DWFTRIG : DWORD;
	BYINBITNO : BYTE;
	BYINBITNOOLD : BYTE;
	XSTATEENTRY : BOOL;
	ETMSTATE_INT : L_TB2P_States := L_TB2P_States.DISABLED;
	ETMSTATE_OLD : L_TB2P_States;
	XFIRSTCYCLE : BOOL := TRUE;
	PBOOL : POINTER TO BOOL;
	PBYTE : POINTER TO BYTE;
	PINT : POINTER TO INT;
	PDINT : POINTER TO DINT;
	PUINT : POINTER TO UINT;
	PSINT : POINTER TO SINT;
	PWORD : POINTER TO WORD;
	PDWORD : POINTER TO DWORD;
	PREAL : POINTER TO REAL;
	PLREAL : POINTER TO LREAL;
	PSTRING : POINTER TO STRING;
	DIFRAME : DINT;
	DIFRAMEPAR : DINT;
	_ESUBCOMPTYPE : UDINT;
	_SLICINFO : STRING(10);
	EXTMODULEHANDLER : L_IMHP_IModuleHandler;
	CHILDMODULEHANDLERINT : L_IMHP_IModuleHandler;
	L_IE1P_SETERROR1 : L_IE1P_SetError := STRUCT(ModuleHandler := ExtModuleHandler);
	_ITFLENZEVENDORIDCHECKER : L_UBUP_IChecker;
	_ITFMCCALLINFOFASSADE : L_UM1P_IMCCallInfo;
	_ITASKIDX : INT;
	_ICALLTASKINDEX : INT;
	_XMULTICOREACTIVE : BOOL;
	MODULEHANDLER : L_IMHP_IModuleHandler;
END_VAR
END_FUNCTION_BLOCK

METHOD CALL_ALLOCPOINTADR
END_METHOD

METHOD CALL_CHECKREQUESTS
END_METHOD

METHOD CALL_ERRORRESETACTIVE
END_METHOD

METHOD CALL_ERRORHANDLER
END_METHOD

METHOD CALL_ERRORHANDLER_SCERRORINFO
END_METHOD

METHOD CALL_FBMETHODS
END_METHOD

METHOD CALL_FIRSTCYCLE
END_METHOD

METHOD CALL_INITDONE
END_METHOD

METHOD CALL_INITROUTINE
END_METHOD

METHOD CALL_INTERNALCTRL
END_METHOD

METHOD CALL_OUTPUT
END_METHOD

METHOD CALL_REQUESTS_EXT
END_METHOD

METHOD CALL_RESETCOMMANDS
END_METHOD

METHOD CALL_RESETOUTPUT
END_METHOD

METHOD CALL_RESETWARNINGS
END_METHOD

METHOD CALL_SETERROR
END_METHOD

METHOD CALL_SYSTEMFAULT : BOOL
END_METHOD

METHOD CALL_TMFUNCTIONALITY
END_METHOD

METHOD INIT_SETERRORFBS
END_METHOD

METHOD HANDLELFASTFRAMEINFORMATION
VAR_INPUT
	CHILDMODULEHANDLE : L_IMHP_IModuleHandler;
	XMODULEACTIVATED : BOOL;
END_VAR
END_METHOD

METHOD SETADDMODULEINFO
VAR_INPUT
	ESUBCOMPTYPE : UDINT;
	SLICINFO : STRING(10);
END_VAR
END_METHOD

METHOD HANDOVERRESOURCE : BOOL
VAR_INPUT
	ITFRESOURCE : L_UBUP_IUnknown;
END_VAR
END_METHOD

METHOD REQUESTINTERFACE : BOOL
VAR_INPUT
	ID : DINT;
	PITFUNKNOWN : POINTER TO L_UBUP_IUnknown;
END_VAR
END_METHOD

METHOD CALL_S000_CYCLIC
END_METHOD

METHOD CALL_S001_INIT
END_METHOD

METHOD CALL_S996_STOP
END_METHOD

METHOD CALL_S999_ERROR
END_METHOD

METHOD CALL_STATEMACHINE
END_METHOD

METHOD CALL_STATEMACHINE_OUT
END_METHOD

METHOD FB_INIT : BOOL
VAR_INPUT
	BINITRETAINS : BOOL;
	BINCOPYCODE : BOOL;
END_VAR
END_METHOD

(* ---- L_TB2P_TM_MOTIONCONTROL.pou ---- *)
FUNCTION_BLOCK L_TB2P_TM_MOTIONCONTROL EXTENDS L_TB2P_TM_Base
VAR_IN_OUT
	AXIS : AXIS_REF;
END_VAR
VAR
	TM_MOTIONCONTROLCONFIG : L_TB2P_ModuleHandlerConfig;
	PINPUTBASE : POINTER TO L_TB2P_BasicMotionBaseIn;
	POUTPUTBASE : POINTER TO L_TB2P_BasicMotionBaseOut;
	XSETHOMEPOSSTATEINDEPENDENTACTIVE : BOOL;
	_PSCPARVISU : POINTER TO L_TB2P_scPar_TM_MotionControl;
	_PSFMOTIONCTRL : POINTER TO L_TB2P_scSF_TM_MotionControl;
	PABCCTRL : POINTER TO L_TB2P_scCtrlBasicMotion;
	XAXISNOTENABLED : BOOL;
	XINVALIDINPUTJOGPOSJOGNEG : BOOL;
	XINTERRUPTHOMINGBYHALT : BOOL;
	FBTEMPLATEABC : L_MC1P_Template;
	PFBTEMPLATEABC : POINTER TO L_MC1P_Template_ForAxis;
	RABC : REFERENCE TO L_MC1P_AxisBasicControl_Internal;
	SCDATAABC : L_MC1P_AxisBasicControlInstanceData;
	PAXISINST : POINTER TO AXIS_REF;
	_XABORTINTERNAL : BOOL;
	_XCALLRESETABORT : BOOL;
	SCABCIN : L_MC1P_AxisBasicControlInput_Internal;
	SCABCOUT : L_MC1P_AxisBasicControlOutput_Internal;
	XSETJERKDEC : BOOL;
	XJOGGINGSETJERKDEC : BOOL;
	HWLIMITSWITCHINTERFACE : L_MC1P_HWLimitSwitchInterface;
	FB_READAXISINFO : MC_ReadAxisInfo;
	XLIMITERCONTROLVALID : BOOL;
	DWLIMITERCONTROL : DWORD;
	XTMSTOP : BOOL;
	XHALT_OLD : BOOL;
	XABORT_OLD : BOOL;
	SCPARMOTIONCONTROL_INT : L_TB2P_scPar_TM_MotionControl;
	XAXISNOTSTANDSTILL : BOOL;
	XAXISISHOMING : BOOL;
	XHOMINGNOTPOSSIBLE : BOOL;
	XAXISNOTHOMED : BOOL;
	XHOMEEXECUTE_OLD : BOOL := FALSE;
	XHALTBUSY_INT : BOOL;
	XHALTDONE_INT : BOOL;
	XHALTDONE_OLD : BOOL;
	XHOMINGBUSY_INT : BOOL;
	XHOMINGDONE_INT : BOOL;
	XJOGGINGBUSY_INT : BOOL;
	XABORTBUSY_INT : BOOL;
	XABORTDONE_INT : BOOL;
	XABORTDONE_OLD : BOOL;
	XQSPAPPLTOSTOP : BOOL;
	XSWITCHTOSTOP : BOOL;
	XDONENEXTCYCLE_INT : BOOL := TRUE;
	XISHOMED_INT : BOOL;
	XDISABLEEXTERNALSTATE_INT : BOOL;
	XMOVEBASICFUNCTION_INT : BOOL;
	XMOVEBASICFUNCTION_OLD : BOOL;
	EABCFUNCSTATE_OLD : L_MC1P_ABC_State;
	XMOVEVELACTIVE_INT : BOOL;
	XMOVERELACTIVE_INT : BOOL;
	XMOVEABSACTIVE_INT : BOOL;
	XQSPACTIVE_INT : BOOL;
	LWTCHECKSUM : LWORD;
	C_IJOGGING : INT := 1;
	LRJERKDEC : LREAL;
	LRJOGGINGJERKDEC : LREAL;
	REMAININGTIMEOFPROFILE : LREAL;
	REMAININGTIMEOFPROFILEAVAILABLE : BOOL;
END_VAR
END_FUNCTION_BLOCK

METHOD CALL_ALLOCPOINTADR
END_METHOD

METHOD CALL_ERRORRESETACTIVE
END_METHOD

METHOD CALL_ERRORHANDLER
END_METHOD

METHOD CALL_ERRORHANDLER_SCERRORINFO
END_METHOD

METHOD CALL_FBMETHODS
END_METHOD

METHOD CALL_INITROUTINE
END_METHOD

METHOD CALL_INTERNALCTRL
END_METHOD

METHOD CALL_MC1P_HWLIMITSWITCH
END_METHOD

METHOD CALL_OUTPUT
END_METHOD

METHOD CALL_REQUESTS_EXT
END_METHOD

METHOD CALL_RESETCOMMANDS
END_METHOD

METHOD CALL_RESETOUTPUT
END_METHOD

METHOD CALL_RESETSETERROR
VAR_IN_OUT
	AXIS : AXIS_REF;
END_VAR
END_METHOD

METHOD CALL_RESETWARNINGS
END_METHOD

METHOD CALL_SETERROR
END_METHOD

METHOD CALL_SYSTEMFAULT : BOOL
END_METHOD

METHOD ABCABORT
END_METHOD

METHOD ABCRESETABORT
END_METHOD

METHOD ABCRESETFINISHPOSITIONING
END_METHOD

METHOD ABCRESETHALT
END_METHOD

METHOD ABCRESETHOMEEXECUTE
END_METHOD

METHOD ABCRESETMOVEABSEXECUTE
END_METHOD

METHOD ABCRESETMOVERELEXECUTE
END_METHOD

METHOD ABCRESETMOVEVELEXECUTE
END_METHOD

METHOD CALL_ABC
END_METHOD

METHOD CALL_ABC_INPUT
END_METHOD

METHOD CALL_ABC_INPUT_PROFILEPARAMETER
END_METHOD

METHOD CALL_MC_READLIMITERWORD
END_METHOD

METHOD CALL_READAXISINFO
END_METHOD

METHOD CALL_S000_CYCLIC_OUT
END_METHOD

METHOD CALL_S003_HOMING_OUT
END_METHOD

METHOD CALL_S009_FINISHPOSITIONING_OUT
END_METHOD

METHOD CALL_S010_JOGGING_OUT
END_METHOD

METHOD CALL_S013_MOVEVEL_OUT
END_METHOD

METHOD CALL_S014_MOVEABS_OUT
END_METHOD

METHOD CALL_S015_MOVEREL_OUT
END_METHOD

METHOD CALL_S017_EXTERNAL_OUT
END_METHOD

METHOD CALL_S996_STOP_OUT
END_METHOD

METHOD CALL_S999_ERROR_OUT
END_METHOD

METHOD CALL_STATEMACHINE_OUT
END_METHOD

METHOD CALL_T000_ALLSTATES_OUT
END_METHOD

METHOD CALL_S000_CYCLIC
END_METHOD

METHOD CALL_S001_INIT
END_METHOD

METHOD CALL_S002_STANDBY
END_METHOD

METHOD CALL_S003_HOMING
END_METHOD

METHOD CALL_S009_FINISHPOSITIONING
END_METHOD

METHOD CALL_S010_JOGGING
END_METHOD

METHOD CALL_S013_MOVEVEL
END_METHOD

METHOD CALL_S014_MOVEABS
END_METHOD

METHOD CALL_S015_MOVEREL
END_METHOD

METHOD CALL_S996_STOP
END_METHOD

METHOD CALL_S999_ERROR
END_METHOD

METHOD CALL_STATEMACHINE
END_METHOD

METHOD CALL_T000_ALLSTATES
END_METHOD

METHOD CALL_T000_CTRLBASICMOTION
END_METHOD

(* ---- L_TB2P_TP_CONVERTER.pou ---- *)
FUNCTION_BLOCK L_TB2P_TP_CONVERTER
VAR_INPUT
	XENABLE : BOOL;
	TPRECDATA : L_MC1P.L_MC1P_TpReceiveData;
	DWTPDELAYACTPOS : DWORD;
	LRTRANSMITCYCLESSETPOS : LREAL;
	XTARGETPOSISSETPOS : BOOL;
	LRCYCPOSTARGET : LREAL;
	LRCYCLELENGTHTARGET : LREAL;
	ETRAVERSINGRANGETARGET : L_MC1P_TraversingRange;
	DICOMPENSATIONVALUE : DINT := 0;
END_VAR
VAR_OUTPUT
	XTPRECEIVED : BOOL;
	LRTPPOSOUT : LREAL;
END_VAR
VAR
	ALRRINGBUFFERPOS : ARRAY [0..20] OF LREAL := [21(0)];
	ALRRINGBUFFERPOSDUMMY : ARRAY [0..20] OF LREAL := [21(0)];
	DWTIMESTAMPDIFF : DWORD;
	DWCYCLES : DWORD;
	DWTIMESTAMPOLD : DWORD;
	DWRESIDUAL : DWORD;
	LRDELTAPOSCYCLE : LREAL;
	LRTASKCYCLE : LREAL;
	DWTASKCYCLE_US : DWORD;
	XINIT : BOOL := FALSE;
	DWTRANSMITTIMESETPOS : DWORD;
	WINITCYCLES : WORD;
END_VAR
END_FUNCTION_BLOCK

METHOD CALL_RINGBUFFER
END_METHOD

(* ---- L_TB2P_VISUPOOL.pou ---- *)
FUNCTION_BLOCK L_TB2P_VISUPOOL
VAR
	M_STNAMESPACE : STRING(80);
	M_STHELPVARID : STRING;
	M_STHELPVARPATH : STRING(255);
	M_STHELP : STRING;
	M_REGISTERIMAGES : BOOL := TRUE;
END_VAR
END_FUNCTION_BLOCK

METHOD FB_INIT : BOOL
VAR_INPUT
	BINITRETAINS : BOOL;
	BINCOPYCODE : BOOL;
END_VAR
END_METHOD

METHOD FB_REINIT : BOOL
END_METHOD

METHOD FB_EXIT : BOOL
VAR_INPUT
	BINCOPYCODE : BOOL;
END_VAR
END_METHOD

(* ---- L_UBUP_REQUESTTRANSITIONEDGECHECKCONDITION.pou ---- *)
FUNCTION_BLOCK L_UBUP_REQUESTTRANSITIONEDGECHECKCONDITION EXTENDS L_UBUP_RequestTransitionEdge
END_FUNCTION_BLOCK

METHOD EDGEUPIMPL : BOOL
END_METHOD
